--- program BumperR_C (robot ABB IRB 1300-10/1.15) ---
  Smooth(1)
  Set speed (1000.0 mm/s)
  Set Ref.: Bumper_R
  Set Tool: Generic Paint Sprayer
  Show Generic Paint Sprayer
  MoveJ 1 to (-1936.32, -807.88, 631.21) mm, rotated rx 93.18 ry 4.14 rz 127.64 deg; joints [-99.533, -17.421, 17.763, 90.671, 92.041, 174.508, 166.076, 424.987, 537.758]
  MoveL 2 to (-1936.32, -807.88, 631.21) mm, rotated rx 93.18 ry 4.14 rz 127.64 deg; joints [-99.533, -17.421, 17.763, 90.671, 92.041, 174.508, 166.076, 424.987, 537.758]
  MoveL 3 to (-1857.02, -747.22, 625.67) mm, rotated rx 93.18 ry 4.14 rz 127.64 deg; joints [-99.533, -17.421, 17.763, 90.671, 92.041, 174.508, 245.383, 485.648, 543.299]
  MoveL 4 to (-1857.02, -747.22, 625.67) mm, rotated rx 93.18 ry 4.14 rz 127.64 deg; joints [-99.533, -17.421, 17.763, 90.671, 92.041, 174.508, 245.383, 485.648, 543.299]
  Set speed (200.0 mm/s)
  MoveL 5 to (-1854.92, -751.4, 608.66) mm, rotated rx 92.71 ry 3.53 rz 127.58 deg; joints [-99.511, -17.421, 17.763, 90.568, 92.041, 175.269, 247.254, 481.589, 561.94]
  MoveL 6 to (-1853.09, -755.07, 592.18) mm, rotated rx 92.47 ry 3.35 rz 126.5 deg; joints [-99.489, -17.145, 17.763, 90.433, 93.086, 175.269, 247.254, 484.938, 580.964]
  MoveL 7 to (-1851.52, -758.47, 576.48) mm, rotated rx 93.66 ry 4.99 rz 126.32 deg; joints [-99.364, -17.145, 16.133, 90.721, 93.228, 174.897, 247.254, 485.358, 580.964]
  MoveL 8 to (-1850.74, -761.61, 561.83) mm, rotated rx 94.86 ry 6.58 rz 126.56 deg; joints [-99.364, -17.392, 14.819, 91.032, 93.106, 174.504, 247.642, 485.358, 580.964]
  MoveL 9 to (-1850.48, -763.96, 548.75) mm, rotated rx 96.79 ry 9.07 rz 127.08 deg; joints [-99.364, -17.665, 14.066, 91.464, 92.867, 172.428, 247.79, 485.358, 580.964]
  MoveL 10 to (-1851.52, -765.27, 536.72) mm, rotated rx 100.03 ry 13.16 rz 127.84 deg; joints [-99.41, -17.665, 13.808, 92.093, 92.867, 167.569, 247.288, 485.542, 580.964]
  MoveL 11 to (-1854.14, -765.79, 525.73) mm, rotated rx 106.46 ry 20.29 rz 130.44 deg; joints [-99.565, -17.69, 13.808, 93.445, 92.604, 158.33, 247.288, 485.542, 571.446]
  MoveL 12 to (-1858.59, -765.01, 515.26) mm, rotated rx 114.08 ry 25.91 rz 135.64 deg; joints [-99.582, -18.538, 13.808, 95.79, 90.846, 150.452, 247.288, 485.542, 548.94]
  MoveL 13 to (-1865.65, -762.91, 505.32) mm, rotated rx 122.27 ry 29.64 rz 141.93 deg; joints [-99.582, -19.151, 13.808, 98.838, 88.998, 143.312, 247.792, 485.542, 521.609]
  MoveL 14 to (-1874.81, -759.25, 495.64) mm, rotated rx 129.05 ry 31.24 rz 147.4 deg; joints [-99.584, -19.274, 13.808, 101.789, 87.65, 137.836, 247.792, 485.542, 499.519]
  MoveL 15 to (-1886.32, -754.02, 486.49) mm, rotated rx 136.02 ry 31.67 rz 153.13 deg; joints [-99.584, -19.274, 13.808, 105.29, 86.453, 132.536, 248.559, 488.116, 473.738]
  MoveL 16 to (-1899.66, -746.96, 478.12) mm, rotated rx 142.32 ry 31.02 rz 158.3 deg; joints [-99.584, -19.274, 13.808, 108.952, 85.547, 127.949, 249.413, 495.397, 447.495]
  MoveL 17 to (-1915.36, -738.32, 470.27) mm, rotated rx 145.68 ry 30.62 rz 160.83 deg; joints [-99.727, -19.274, 13.808, 110.865, 85.547, 125.497, 241.966, 507.62, 437.97]
  MoveL 18 to (-1931.84, -728.38, 462.94) mm, rotated rx 149.65 ry 30.54 rz 163.43 deg; joints [-99.727, -19.274, 13.808, 112.679, 85.974, 122.436, 231.514, 526.497, 429.039]
  MoveL 19 to (-1948.58, -717.13, 456.14) mm, rotated rx 152.24 ry 30.71 rz 164.95 deg; joints [-99.727, -19.274, 13.808, 113.594, 86.536, 120.405, 217.15, 545.852, 427.786]
  MoveL 20 to (-1964.28, -704.84, 450.12) mm, rotated rx 153.43 ry 32.04 rz 165.14 deg; joints [-99.727, -19.274, 12.548, 112.864, 87.093, 120.405, 195.765, 569.427, 430.366]
  MoveL 21 to (-1978.14, -692.28, 444.63) mm, rotated rx 153.62 ry 34.41 rz 164.34 deg; joints [-99.727, -19.274, 11.863, 110.908, 88.335, 120.405, 170.573, 593.858, 448.118]
  MoveL 22 to (-1990.18, -678.94, 439.66) mm, rotated rx 153.89 ry 36.46 rz 163.77 deg; joints [-99.727, -19.274, 11.132, 109.278, 89.362, 120.405, 149.601, 617.715, 462.665]
  MoveL 23 to (-2001.17, -663.76, 435.73) mm, rotated rx 154.97 ry 37.74 rz 164.05 deg; joints [-99.727, -19.274, 9.965, 108.565, 89.866, 120.405, 133.981, 642.57, 464.996]
  MoveL 24 to (-2011.11, -646.76, 432.33) mm, rotated rx 155.17 ry 39.62 rz 163.56 deg; joints [-99.727, -19.274, 9.284, 107.066, 90.789, 120.405, 116.666, 668.628, 477.923]
  MoveL 25 to (-2020.53, -627.4, 429.98) mm, rotated rx 157.04 ry 40.04 rz 164.76 deg; joints [-99.727, -19.274, 9.179, 107.28, 91.159, 119.081, 107.159, 693.484, 477.923]
  MoveL 26 to (-2029.16, -606.21, 428.41) mm, rotated rx 158.94 ry 40.39 rz 165.99 deg; joints [-99.727, -19.274, 9.179, 107.517, 91.545, 117.663, 98.62, 719.886, 477.702]
  MoveL 27 to (-2037.01, -583.97, 427.36) mm, rotated rx 160.23 ry 41.22 rz 166.67 deg; joints [-99.727, -19.274, 8.49, 107.168, 91.913, 117.224, 88.381, 748.859, 477.702]
  MoveL 28 to (-2044.59, -558.86, 426.58) mm, rotated rx 161.39 ry 42.2 rz 167.25 deg; joints [-99.727, -19.274, 7.571, 106.639, 92.277, 117.063, 77.677, 781.257, 477.702]
  MoveL 29 to (-2052.44, -527.72, 426.05) mm, rotated rx 163.85 ry 43.54 rz 168.72 deg; joints [-99.727, -19.274, 6.547, 106.072, 92.915, 116.051, 66.17, 823.308, 477.702]
  MoveL 30 to (-2059.77, -491.62, 425.27) mm, rotated rx 165.59 ry 45.05 rz 169.7 deg; joints [-99.727, -19.274, 4.995, 105.182, 93.397, 116.035, 54.117, 870.014, 477.702]
  MoveL 31 to (-2066.57, -450.02, 425.01) mm, rotated rx 167.57 ry 45.52 rz 171.06 deg; joints [-99.727, -19.274, 4.773, 105.136, 93.752, 114.842, 46.502, 916.944, 477.702]
  MoveL 32 to (-2072.32, -407.9, 424.48) mm, rotated rx 169.72 ry 45.69 rz 172.6 deg; joints [-99.727, -19.274, 4.772, 105.319, 94.067, 113.385, 40.863, 963.663, 477.247]
  MoveL 33 to (-2076.77, -369.45, 424.48) mm, rotated rx 172.37 ry 44.66 rz 174.62 deg; joints [-99.739, -19.073, 4.773, 106.624, 94.061, 111.6, 40.863, 1004.094, 466.401]
  MoveL 34 to (-2080.43, -332.3, 424.22) mm, rotated rx 173.02 ry 44.75 rz 175.07 deg; joints [-99.739, -19.073, 4.699, 106.632, 94.169, 111.22, 37.023, 1042.993, 466.401]
  MoveL 35 to (-2083.57, -293.84, 424.22) mm, rotated rx 174.33 ry 44.89 rz 175.99 deg; joints [-99.739, -19.073, 4.643, 106.655, 94.406, 110.368, 33.624, 1084.71, 466.401]
  MoveL 36 to (-2086.45, -254.34, 423.96) mm, rotated rx 174.99 ry 44.96 rz 176.45 deg; joints [-99.739, -19.073, 4.578, 106.671, 94.512, 109.977, 30.611, 1125.93, 466.401]
  MoveL 37 to (-2088.81, -213.79, 423.96) mm, rotated rx 174.99 ry 44.96 rz 176.45 deg; joints [-99.739, -19.073, 4.578, 106.671, 94.512, 109.977, 28.256, 1166.48, 466.401]
  MoveL 38 to (-2090.9, -172.19, 423.96) mm, rotated rx 176.32 ry 45.06 rz 177.39 deg; joints [-99.739, -19.073, 4.541, 106.71, 94.746, 109.105, 25.989, 1211.272, 466.401]
  MoveL 39 to (-2092.47, -129.81, 423.96) mm, rotated rx 177.06 ry 44.63 rz 177.93 deg; joints [-99.74, -19.032, 4.541, 107.175, 94.739, 108.614, 25.988, 1254.666, 462.512]
  MoveL 40 to (-2093.78, -86.9, 424.22) mm, rotated rx 178.13 ry 43.73 rz 178.71 deg; joints [-99.74, -19.032, 4.541, 108.117, 94.642, 107.976, 27.818, 1299.855, 454.042]
  MoveL 41 to (-2094.82, -43.48, 424.22) mm, rotated rx 179.06 ry 43.76 rz 179.35 deg; joints [-99.74, -19.032, 4.528, 108.161, 94.823, 107.343, 26.715, 1345.663, 454.042]
  MoveL 42 to (-2095.87, -0.05, 424.22) mm, rotated rx -180 ry 43.76 rz -180 deg; joints [-99.74, -19.031, 4.528, 108.215, 95.004, 106.699, 25.661, 1391.44, 454.042]
  MoveL 43 to (-2094.82, 43.64, 424.22) mm, rotated rx -179.06 ry 43.76 rz -179.35 deg; joints [-99.572, -19.031, 4.528, 108.223, 95.03, 106.004, 25.661, 1437.299, 454.038]
  MoveL 44 to (-2093.78, 87.07, 424.22) mm, rotated rx -178.13 ry 43.73 rz -178.71 deg; joints [-99.397, -19.031, 4.528, 108.24, 95.047, 105.308, 25.661, 1482.893, 453.951]
  MoveL 45 to (-2092.47, 129.97, 423.96) mm, rotated rx -177.06 ry 44.63 rz -177.93 deg; joints [-99.397, -19.031, 3.701, 107.472, 95.232, 105.308, 23.483, 1530.189, 456.644]
  MoveL 46 to (-2090.9, 172.35, 423.96) mm, rotated rx -176.32 ry 45.06 rz -177.39 deg; joints [-99.397, -19.031, 3.152, 107.121, 95.314, 105.308, 23.335, 1575.521, 456.873]
  MoveL 47 to (-2088.81, 213.69, 423.96) mm, rotated rx -174.99 ry 44.96 rz -176.45 deg; joints [-99.155, -19.031, 3.152, 107.158, 95.314, 104.338, 24.086, 1619.712, 456.608]
  MoveL 48 to (-2086.45, 254.24, 423.96) mm, rotated rx -174.99 ry 44.96 rz -176.45 deg; joints [-99.155, -19.031, 3.152, 107.158, 95.314, 104.338, 26.44, 1660.262, 456.608]
  MoveL 49 to (-2083.57, 293.74, 424.22) mm, rotated rx -174.33 ry 44.89 rz -175.99 deg; joints [-99.036, -19.031, 3.152, 107.184, 95.314, 103.855, 28.685, 1701.202, 456.156]
  MoveL 50 to (-2080.43, 332.2, 424.22) mm, rotated rx -173.02 ry 44.75 rz -175.07 deg; joints [-98.796, -19.031, 3.152, 107.239, 95.314, 102.892, 30.574, 1742.548, 455.762]
  MoveL 51 to (-2076.77, 369.61, 424.48) mm, rotated rx -172.55 ry 44.21 rz -174.79 deg; joints [-98.796, -19.031, 3.152, 107.761, 95.299, 102.576, 35.936, 1781.615, 451.106]
  MoveL 52 to (-2072.32, 408.07, 424.48) mm, rotated rx -169.84 ry 45.47 rz -172.72 deg; joints [-98.796, -19.031, 1.231, 106.589, 95.496, 102.576, 34.759, 1829.747, 451.505]
  MoveL 53 to (-2066.57, 450.19, 425.01) mm, rotated rx -167.57 ry 45.52 rz -171.06 deg; joints [-98.445, -19.031, 0.86, 106.319, 95.496, 101.296, 37.362, 1877.139, 451.505]
  MoveL 54 to (-2059.77, 491.52, 425.27) mm, rotated rx -165.59 ry 45.05 rz -169.7 deg; joints [-98.116, -19.031, 0.86, 106.5, 95.496, 99.832, 42.872, 1922.962, 449.946]
  MoveL 55 to (-2052.44, 527.89, 426.05) mm, rotated rx -164.03 ry 43.34 rz -168.89 deg; joints [-97.985, -19.031, 0.86, 107.995, 95.496, 98.569, 54.252, 1966.24, 436.98]
  MoveL 56 to (-2044.59, 558.76, 426.58) mm, rotated rx -161.39 ry 42.2 rz -167.25 deg; joints [-97.449, -19.031, 0.86, 108.62, 95.496, 96.434, 61.329, 2005.2, 431.733]
  MoveL 57 to (-2037.01, 584.14, 427.36) mm, rotated rx -159.73 ry 41 rz -166.38 deg; joints [-97.078, -19.031, 0.86, 109.449, 95.496, 94.99, 69.884, 2037.373, 424.494]
  MoveL 58 to (-2029.16, 606.11, 428.41) mm, rotated rx -158.46 ry 40.17 rz -165.72 deg; joints [-96.751, -19.031, 0.86, 109.96, 95.496, 93.867, 77.91, 2064.498, 419.566]
  MoveL 59 to (-2020.53, 627.3, 429.98) mm, rotated rx -157.04 ry 40.04 rz -164.76 deg; joints [-96.751, -19.031, 0.73, 109.835, 95.79, 92.944, 85.922, 2089.517, 419.566]
  MoveL 60 to (-2011.11, 646.92, 432.33) mm, rotated rx -155.42 ry 39.47 rz -163.79 deg; joints [-96.299, -19.031, 0.73, 109.921, 95.79, 91.528, 93.399, 2114.204, 416.903]
  MoveL 61 to (-2001.17, 663.93, 435.73) mm, rotated rx -155.23 ry 37.59 rz -164.28 deg; joints [-96.106, -19.031, 0.73, 111.729, 95.79, 91.025, 109.339, 2138.748, 399.131]
  MoveL 62 to (-1990.18, 678.84, 439.66) mm, rotated rx -154.15 ry 36.32 rz -163.99 deg; joints [-95.651, -19.031, 0.73, 112.633, 95.79, 89.863, 121.839, 2160.968, 388.385]
  MoveL 63 to (-1978.14, 692.44, 444.63) mm, rotated rx -153.62 ry 34.41 rz -164.34 deg; joints [-95.237, -19.031, 0.73, 114.331, 95.79, 89.028, 139.219, 2183.618, 370.37]
  MoveL 64 to (-1964.28, 705, 450.12) mm, rotated rx -153.68 ry 31.92 rz -165.34 deg; joints [-94.887, -19.031, 0.73, 116.823, 95.79, 88.593, 162.975, 2206.59, 345.904]
  MoveL 65 to (-1948.58, 717.03, 456.14) mm, rotated rx -152.24 ry 30.71 rz -164.95 deg; joints [-94.076, -19.031, 0.73, 117.431, 95.79, 86.979, 178.162, 2227.857, 335.852]
  MoveL 66 to (-1931.84, 728.28, 462.94) mm, rotated rx -149.65 ry 30.54 rz -163.43 deg; joints [-94.076, -19.031, 0.546, 116.895, 96.626, 85.113, 192.486, 2247.762, 335.852]
  MoveL 67 to (-1915.36, 738.49, 470.27) mm, rotated rx -145.68 ry 30.62 rz -160.83 deg; joints [-94.076, -19.031, -0.772, 115.634, 97.273, 83.206, 202.648, 2270.964, 335.852]
  MoveL 68 to (-1899.66, 747.12, 478.12) mm, rotated rx -142.32 ry 31.02 rz -158.3 deg; joints [-94.076, -19.031, -2.193, 114.066, 97.487, 81.93, 210.701, 2287.64, 335.852]
  MoveL 69 to (-1886.32, 753.92, 486.49) mm, rotated rx -136.33 ry 31.66 rz -153.39 deg; joints [-94.433, -19.031, -5.824, 111.213, 97.484, 80.878, 211.61, 2307.705, 336.675]
  MoveL 70 to (-1874.81, 759.15, 495.64) mm, rotated rx -129.05 ry 31.24 rz -147.4 deg; joints [-94.884, -19.031, -10.183, 108.228, 97.484, 79.328, 211.337, 2327.777, 336.675]
  MoveL 71 to (-1865.65, 762.82, 505.32) mm, rotated rx -121.95 ry 29.53 rz -141.67 deg; joints [-95.215, -19.031, -14.028, 105.588, 97.484, 76.903, 210.999, 2343.299, 336.676]
  MoveL 72 to (-1858.59, 764.91, 515.26) mm, rotated rx -113.78 ry 25.73 rz -135.42 deg; joints [-95.671, -19.031, -18.384, 102.957, 97.484, 73.021, 209.766, 2357.906, 336.68]
  MoveL 73 to (-1854.14, 765.7, 525.73) mm, rotated rx -105.9 ry 19.78 rz -130.1 deg; joints [-96.122, -19.031, -22.104, 100.789, 97.484, 67.188, 208.374, 2368.079, 336.681]
  MoveL 74 to (-1851.52, 765.43, 536.72) mm, rotated rx -100.03 ry 13.16 rz -127.84 deg; joints [-96.122, -19.031, -23.565, 99.944, 97.888, 59.882, 208.876, 2376.573, 336.681]
  MoveL 75 to (-1850.48, 763.86, 548.75) mm, rotated rx -97.28 ry 9.68 rz -127.23 deg; joints [-96.122, -19.033, -23.565, 99.613, 98.284, 55.461, 209.792, 2376.573, 333.147]
  MoveL 76 to (-1850.74, 761.51, 561.83) mm, rotated rx -94.38 ry 5.95 rz -126.45 deg; joints [-96.122, -19.324, -23.565, 99.024, 98.427, 50.977, 208.321, 2376.573, 329.103]
  MoveL 77 to (-1851.52, 758.63, 576.48) mm, rotated rx -93.66 ry 4.99 rz -126.32 deg; joints [-96.122, -19.541, -23.565, 98.92, 98.45, 49.99, 207.062, 2376.573, 316.404]
  MoveL 78 to (-1853.09, 755.23, 592.18) mm, rotated rx -92.47 ry 3.35 rz -126.5 deg; joints [-96.122, -19.581, -23.565, 98.982, 98.785, 48.026, 205.933, 2376.573, 304.255]
  MoveL 79 to (-1854.92, 751.31, 608.66) mm, rotated rx -92.71 ry 3.53 rz -127.58 deg; joints [-95.902, -19.193, -23.565, 99.595, 99.379, 48.025, 205.932, 2376.585, 287.089]
  MoveL 80 to (-1857.02, 747.38, 625.67) mm, rotated rx -92.47 ry 3.22 rz -127.55 deg; joints [-95.903, -19.46, -23.565, 99.595, 99.364, 47.903, 203.405, 2376.585, 270.462]
  Set speed (1000.0 mm/s)
  MoveL 81 to (-1857.02, 747.38, 625.67) mm, rotated rx -92.47 ry 3.22 rz -127.55 deg; joints [-95.903, -19.46, -23.565, 99.595, 99.364, 47.903, 203.405, 2376.585, 270.462]
  MoveL 82 to (-1936.37, 808.08, 629.98) mm, rotated rx -92.47 ry 3.22 rz -127.55 deg; joints [-95.903, -19.46, -23.565, 99.595, 99.364, 47.903, 124.049, 2437.282, 266.151]
  Set speed (1000.0 mm/s)
  MoveL 83 to (-1866.33, 853.74, 600.09) mm, rotated rx -83.63 ry -41.53 rz -164.5 deg; joints [-62.31, -26.599, -19.684, 114.622, 92.23, 9.806, 295.721, 2881.383, 207.551]
  MoveL 84 to (-1832.69, 759.94, 608.4) mm, rotated rx -85.23 ry -1.7 rz -160.41 deg; joints [0, -20.746, 0, 63.366, 46.167, 29.285, 22.945, 2896.284, 466.116]
  MoveL 85 to (-1832.69, 759.94, 608.4) mm, rotated rx -85.23 ry -1.7 rz -160.41 deg; joints [0, -20.746, 0, 63.366, 46.167, 29.285, 22.945, 2896.284, 466.116]
  Set speed (200.0 mm/s)
  MoveL 86 to (-1807.05, 769.62, 608.4) mm, rotated rx -85.47 ry -1.55 rz -161.18 deg; joints [0.673, -20.681, 0, 63.662, 46.168, 29.285, 53.093, 2915.113, 464.886]
  MoveL 87 to (-1774.35, 780.87, 608.4) mm, rotated rx -86.88 ry -1.04 rz -161.54 deg; joints [0.494, -20.669, 0, 65.263, 46.167, 29.285, 88.293, 2928.573, 454.825]
  MoveL 88 to (-1737.72, 792.64, 608.92) mm, rotated rx -87.13 ry -0.81 rz -164.2 deg; joints [2.732, -20.666, 0, 65.706, 46.49, 29.285, 144.085, 2970.228, 453.078]
  MoveL 89 to (-1699.52, 803.37, 611.02) mm, rotated rx -87.04 ry -0.78 rz -165.26 deg; joints [3.621, -20.666, 0, 65.706, 46.681, 29.257, 190.209, 2992.448, 451.942]
  MoveL 90 to (-1699.52, 803.37, 611.02) mm, rotated rx -87.81 ry -2 rz -137.59 deg; joints [-23.141, -21.64, 0, 65.706, 45.639, 29.257, 72.494, 2638.724, 437.476]
  MoveL 91 to (-1692.72, 808.6, 595.58) mm, rotated rx -87.36 ry -2.41 rz -137.69 deg; joints [-23.141, -21.452, 0, 65.706, 45.726, 28.553, 77.414, 2643.64, 455.753]
  MoveL 92 to (-1682.78, 815.66, 576.22) mm, rotated rx -85.22 ry -4.18 rz -138.93 deg; joints [-23.14, -21.036, 0, 65.706, 46.944, 25.645, 86.714, 2657.383, 487.623]
  MoveL 93 to (-1678.33, 821.16, 555.29) mm, rotated rx -92.02 ry 1.97 rz -135.8 deg; joints [-23.14, -21.586, 0, 66.424, 43.225, 34.246, 86.714, 2640.571, 472.908]
  MoveL 94 to (-1642.49, 837.12, 523.37) mm, rotated rx -77.29 ry -8.01 rz -148.28 deg; joints [-23.14, -19.929, 0, 66.424, 55.746, 16.427, 152.9, 2736.554, 595.298]
  MoveL 95 to (-1620.52, 847.58, 496.95) mm, rotated rx -79.58 ry -7.51 rz -144.62 deg; joints [-23.14, -19.686, 0, 66.424, 52.076, 18.199, 155.26, 2721.165, 605.579]
  MoveL 96 to (-1620.52, 847.58, 496.95) mm, rotated rx -99.89 ry 2.5 rz -165.96 deg; joints [-23.14, -12.952, 0, 92.6, 67.432, 18.199, 210.874, 2845.232, 499.77]
  MoveL 97 to (-1641.45, 845.49, 477.07) mm, rotated rx -98.6 ry 2.33 rz -164.94 deg; joints [-23.14, -13.332, 0, 91.157, 66.772, 18.199, 186.996, 2840.685, 528.15]
  MoveL 98 to (-1660.28, 843.13, 455.62) mm, rotated rx -97.18 ry 2.02 rz -164.37 deg; joints [-23.141, -13.834, 0, 89.716, 66.592, 18.199, 170.028, 2839.081, 558.046]
  MoveL 99 to (-1678.33, 840.52, 432.86) mm, rotated rx -96.24 ry 1.87 rz -163.38 deg; joints [-23.141, -14.087, 0, 88.595, 65.882, 18.199, 147.906, 2832.55, 587.081]
  MoveL 100 to (-1695.08, 837.64, 409.05) mm, rotated rx -95.06 ry 1.57 rz -162.84 deg; joints [-23.141, -14.51, 0, 87.369, 65.678, 18.199, 132.362, 2829.437, 617.84]
  MoveL 101 to (-1709.73, 835.02, 384.98) mm, rotated rx -93.88 ry 1.24 rz -162.32 deg; joints [-23.141, -14.941, 0, 86.142, 65.486, 18.199, 119.084, 2826.443, 648.781]
  MoveL 102 to (-1722.28, 832.41, 361.44) mm, rotated rx -92.94 ry 0.99 rz -161.35 deg; joints [-23.141, -15.215, 0, 85.008, 64.801, 18.199, 102.986, 2819.412, 678.238]
  MoveL 103 to (-1732.23, 830.05, 338.68) mm, rotated rx -92 ry 0.68 rz -161.32 deg; joints [-23.127, -15.625, 0, 84.119, 65.017, 18.199, 97.559, 2819.356, 706.065]
  MoveL 104 to (-1740.6, 827.96, 316.96) mm, rotated rx -91.53 ry 0.52 rz -161.31 deg; joints [-23.126, -15.833, 0, 83.678, 65.137, 18.199, 91.508, 2818.353, 730.315]
  MoveL 105 to (-1747.4, 826.13, 295.51) mm, rotated rx -91.06 ry 0.37 rz -160.6 deg; joints [-23.4, -15.978, 0, 83.118, 64.841, 18.199, 82.237, 2810.955, 754.634]
  Set speed (1000.0 mm/s)
  MoveL 106 to (-1747.4, 826.13, 295.51) mm, rotated rx -91.06 ry 0.37 rz -160.6 deg; joints [-23.4, -15.978, 0, 83.118, 64.841, 18.199, 82.237, 2810.955, 754.634]
  MoveL 107 to (-1780.63, 920.43, 297.36) mm, rotated rx -91.06 ry 0.37 rz -160.6 deg; joints [-23.4, -15.978, 0, 83.118, 64.841, 18.199, 49.007, 2905.255, 752.786]
  Set speed (1000.0 mm/s)
  MoveL 108 to (-1840, 893.27, 313.81) mm, rotated rx -106.34 ry 6.01 rz -160.35 deg; joints [-23.4, -17.541, 0, 92.672, 59.812, 27.622, 0.008, 2861.075, 623.578]
  MoveL 109 to (-1804.95, 803.89, 285.83) mm, rotated rx -106.34 ry 6.01 rz -160.35 deg; joints [-23.4, -17.541, 0, 92.672, 59.812, 27.622, 35.053, 2771.694, 651.559]
  MoveL 110 to (-1804.95, 803.89, 285.83) mm, rotated rx -106.34 ry 6.01 rz -160.35 deg; joints [-23.4, -17.541, 0, 92.672, 59.812, 27.622, 35.053, 2771.694, 651.559]
  Set speed (200.0 mm/s)
  MoveL 111 to (-1832.95, 791.59, 290.54) mm, rotated rx -106.49 ry 6.19 rz -159.99 deg; joints [-23.4, -17.541, 0.133, 92.672, 59.412, 27.666, 4.112, 2756.326, 647.26]
  MoveL 112 to (-1858.06, 779.82, 294.2) mm, rotated rx -106.41 ry 7.21 rz -156.92 deg; joints [-26.51, -20.886, 1.667, 90.881, 59.412, 30.95, 0, 2721.012, 647.26]
  MoveL 113 to (-1879.78, 768.57, 296.56) mm, rotated rx -105.99 ry 7.97 rz -154.18 deg; joints [-29.001, -23.988, 2.357, 88.525, 59.412, 34.604, 0, 2695.317, 647.26]
  MoveL 114 to (-1896.78, 758.89, 298.13) mm, rotated rx -106.1 ry 9.48 rz -150.31 deg; joints [-32.699, -26.95, 2.767, 86.07, 59.412, 39.328, 0, 2657.479, 647.26]
  MoveL 115 to (-1911.69, 749.48, 299.17) mm, rotated rx -106.56 ry 10.61 rz -148.24 deg; joints [-34.777, -29.185, 3.342, 84.726, 59.412, 42.61, 0, 2636.415, 647.26]
  MoveL 116 to (-1927.13, 738.75, 299.96) mm, rotated rx -105.67 ry 11.02 rz -145.73 deg; joints [-36.306, -31.519, 3.342, 81.953, 59.412, 45.771, 0, 2619.867, 652.638]
  MoveL 117 to (-1942.56, 726.98, 301) mm, rotated rx -105.75 ry 12.18 rz -143.21 deg; joints [-38.217, -33.858, 3.342, 79.586, 59.412, 49.888, 0, 2598.73, 654.329]
  MoveL 118 to (-1957.74, 714.42, 301.79) mm, rotated rx -105.83 ry 13.67 rz -140.19 deg; joints [-40.307, -36.353, 3.342, 76.719, 59.412, 54.629, 0, 2574.299, 659.016]
  MoveL 119 to (-1971.86, 701.08, 302.57) mm, rotated rx -105.19 ry 14.87 rz -136.61 deg; joints [-42.079, -38.903, 3.342, 72.981, 59.412, 59.147, 0, 2548.829, 669.678]
  MoveL 120 to (-1984.68, 686.95, 303.1) mm, rotated rx -104.58 ry 16.89 rz -131.85 deg; joints [-44.246, -41.542, 3.342, 68.194, 59.412, 64.909, 0, 2512.396, 685.44]
  MoveL 121 to (-1996.19, 672.3, 303.62) mm, rotated rx -105.37 ry 20.17 rz -128.56 deg; joints [-45.598, -43.63, 3.342, 64.184, 59.412, 71.634, 0, 2480.166, 696.443]
  MoveL 122 to (-2006.4, 656.6, 303.88) mm, rotated rx -105.16 ry 23.11 rz -124.63 deg; joints [-46.174, -45.488, 3.342, 58.938, 59.412, 77.967, 0, 2443.432, 714.605]
  MoveL 123 to (-2015.55, 640.12, 304.14) mm, rotated rx -105.39 ry 26.98 rz -121.25 deg; joints [-46.174, -47.75, 3.343, 53.282, 60.14, 85.802, 7.235, 2413.258, 735.61]
  MoveL 124 to (-2023.66, 622.59, 304.14) mm, rotated rx -105.02 ry 30.09 rz -118.16 deg; joints [-46.174, -47.998, 3.343, 49.217, 60.37, 90.526, 0.63, 2370.196, 753.089]
  MoveL 125 to (-2030.47, 604.8, 304.14) mm, rotated rx -104.12 ry 31.18 rz -115.91 deg; joints [-46.181, -48.648, 3.343, 46.493, 60.949, 92.894, 0.01, 2341.413, 766.26]
  MoveL 126 to (-2036.48, 586.75, 303.88) mm, rotated rx -103.81 ry 32.8 rz -114.41 deg; joints [-46.851, -49.255, 3.343, 45.076, 62.033, 95.231, 0, 2316.688, 777.689]
  MoveL 127 to (-2041.98, 569.22, 303.88) mm, rotated rx -105.4 ry 36.74 rz -114.72 deg; joints [-46.853, -49.837, 3.343, 44.146, 63.26, 100.087, 0, 2300.801, 786.26]
  MoveL 128 to (-2046.42, 552.48, 303.62) mm, rotated rx -106.11 ry 42.57 rz -113.12 deg; joints [-47.479, -50.038, 3.343, 41.986, 65.443, 106.494, 0, 2270.786, 809.046]
  MoveL 129 to (-2050.61, 534.69, 303.62) mm, rotated rx -109.1 ry 48.54 rz -114.8 deg; joints [-47.479, -50.429, 3.343, 41.714, 67.353, 112.969, 0, 2258.639, 820.752]
  MoveL 130 to (-2054.53, 514.02, 303.36) mm, rotated rx -110.56 ry 52.74 rz -115.23 deg; joints [-47.479, -50.69, 3.343, 40.989, 68.994, 117.465, 0, 2238.905, 834.382]
  MoveL 131 to (-2058.2, 490.48, 303.88) mm, rotated rx -114 ry 59.08 rz -117.43 deg; joints [-47.479, -50.872, 3.343, 40.753, 71.292, 123.95, 0, 2220.446, 850.258]
  MoveL 132 to (-2061.08, 464.84, 305.97) mm, rotated rx -122.64 ry 66.68 rz -124.9 deg; joints [-47.479, -51.083, 3.343, 41.781, 73.743, 131.949, 0, 2208.96, 860.36]
  MoveL 133 to (-2062.65, 439.2, 310.16) mm, rotated rx -130.58 ry 72.26 rz -131.97 deg; joints [-47.479, -50.951, 3.343, 42.168, 75.885, 137.566, 0.014, 2190.405, 870.985]
  MoveL 134 to (-2062.91, 416.18, 317.48) mm, rotated rx -143.56 ry 74.86 rz -144.52 deg; joints [-47.479, -51.111, 3.343, 43.565, 76.5, 141.58, 0.003, 2178.849, 861.295]
  MoveL 135 to (-2061.86, 396.56, 326.64) mm, rotated rx -154.06 ry 77.62 rz -154.59 deg; joints [-47.479, -50.7, 3.343, 43.858, 77.758, 144.603, 0.003, 2161.713, 861.88]
  MoveL 136 to (-2060.55, 380.6, 335.8) mm, rotated rx 150.62 ry 75.7 rz 151.38 deg; joints [-45.847, -50.793, 3.343, 46.572, 77.758, 156.331, 0, 2171.642, 840.226]
  MoveL 137 to (-2058.72, 368.04, 344.43) mm, rotated rx 152.54 ry 74.9 rz 153.36 deg; joints [-45.847, -50.981, 3.343, 46.912, 77.016, 156.331, 1.624, 2159.565, 823.551]
  MoveL 138 to (-2058.72, 368.04, 344.43) mm, rotated rx 92.19 ry 15.16 rz 98.34 deg; joints [-44.513, -50.981, 6.874, 68.618, 77.016, 213.54, 0.029, 2281.819, 776.099]
  MoveL 139 to (-2057.15, 355.75, 333.7) mm, rotated rx 92.56 ry 14.93 rz 99.84 deg; joints [-45.621, -51.277, 6.873, 68.618, 76.619, 213.86, 0.028, 2259.663, 783.809]
  MoveL 140 to (-2055.32, 342.93, 324.29) mm, rotated rx 92.93 ry 15.77 rz 100.68 deg; joints [-45.895, -51.277, 6.089, 67.95, 76.619, 213.86, 3.03, 2242.747, 789.664]
  MoveL 141 to (-2053.23, 328.54, 316.96) mm, rotated rx 95.76 ry 28.51 rz 101.93 deg; joints [-45.895, -51.277, 6.089, 63.921, 78.506, 202.475, 4.666, 2215.059, 824.396]
  MoveL 142 to (-2051.13, 313.1, 310.68) mm, rotated rx 118.95 ry 67.19 rz 120.96 deg; joints [-45.895, -51.277, 6.033, 50.461, 78.558, 166.142, 4.666, 2125.247, 882.217]
  MoveL 143 to (-2051.92, 299.5, 309.11) mm, rotated rx -151.61 ry 73.09 rz -152.65 deg; joints [-47.318, -58.551, 5.026, 44.393, 78.558, 146.287, 59.413, 2125.246, 882.217]
  MoveL 144 to (-2052.7, 288.51, 308.07) mm, rotated rx -151.22 ry 73.16 rz -152.27 deg; joints [-47.318, -58.551, 4.959, 44.303, 78.693, 146.287, 59.104, 2114.315, 884.068]
  MoveL 145 to (-2053.49, 274.38, 306.76) mm, rotated rx -150.44 ry 73.3 rz -151.48 deg; joints [-47.318, -58.551, 4.866, 44.129, 78.934, 146.254, 59.104, 2100.102, 887.137]
  MoveL 146 to (-2054.27, 258.16, 305.97) mm, rotated rx -149.06 ry 72.23 rz -150.28 deg; joints [-47.226, -59.65, 4.866, 44.129, 78.934, 146.178, 65.904, 2092.744, 886.105]
  MoveL 147 to (-2055.06, 239.33, 305.45) mm, rotated rx -154.8 ry 72.39 rz -155.84 deg; joints [-47.225, -59.873, 4.866, 44.801, 78.77, 147.78, 65.904, 2079.049, 882.098]
  MoveL 148 to (-2056.1, 217.35, 304.93) mm, rotated rx -154.8 ry 72.39 rz -155.84 deg; joints [-47.225, -59.873, 4.866, 44.801, 78.77, 147.78, 64.858, 2057.074, 882.621]
  MoveL 149 to (-2057.15, 191.19, 304.67) mm, rotated rx -160.37 ry 72.86 rz -161.18 deg; joints [-47.225, -59.873, 4.866, 45.256, 78.83, 149.358, 63.555, 2033.518, 881.475]
  MoveL 150 to (-2057.94, 160.84, 304.4) mm, rotated rx -161.41 ry 72.47 rz -162.22 deg; joints [-47.225, -60.055, 4.866, 45.508, 78.575, 149.604, 63.555, 2005.37, 878.309]
  MoveL 151 to (-2058.98, 125, 304.14) mm, rotated rx -165.69 ry 73.35 rz -166.27 deg; joints [-47.225, -60.055, 4.866, 45.553, 79.185, 151.005, 63.203, 1971.107, 883.479]
  MoveL 152 to (-2060.03, 85.5, 303.62) mm, rotated rx -171.28 ry 73.69 rz -171.62 deg; joints [-47.225, -60.055, 4.866, 45.887, 79.393, 152.515, 62.195, 1933.866, 884.39]
  MoveL 153 to (-2060.81, 43.38, 303.36) mm, rotated rx -171.76 ry 73.23 rz -172.11 deg; joints [-47.225, -60.238, 4.866, 46.098, 79.111, 152.676, 62.196, 1893.577, 881.184]
  MoveL 154 to (-2061.6, -0.05, 302.83) mm, rotated rx -180 ry 73.41 rz -180 deg; joints [-47.225, -60.238, 4.866, 46.593, 79.366, 154.887, 61.429, 1853.309, 881.898]
  MoveL 155 to (-2060.81, -43.48, 303.36) mm, rotated rx 171.76 ry 73.23 rz 172.11 deg; joints [-47.225, -60.238, 5.04, 47.132, 79.458, 156.967, 61.428, 1812.212, 881.819]
  MoveL 156 to (-2060.03, -85.6, 303.62) mm, rotated rx 171.28 ry 73.69 rz 171.62 deg; joints [-47.225, -60.101, 5.04, 46.98, 79.805, 156.967, 61.793, 1769.226, 885.263]
  MoveL 157 to (-2058.98, -125.1, 304.14) mm, rotated rx 165.69 ry 73.35 rz 166.27 deg; joints [-47.225, -60.101, 5.219, 47.378, 79.805, 158.339, 62.013, 1731.134, 885.013]
  MoveL 158 to (-2057.94, -160.68, 304.4) mm, rotated rx 161.41 ry 72.47 rz 162.22 deg; joints [-47.225, -60.101, 5.219, 47.887, 79.452, 159.658, 62.365, 1697.132, 879.843]
  MoveL 159 to (-2057.15, -191.29, 304.67) mm, rotated rx 160.37 ry 72.86 rz 161.18 deg; joints [-47.226, -59.919, 5.219, 47.785, 79.783, 159.711, 62.365, 1665.648, 883.012]
  MoveL 160 to (-2056.1, -217.19, 304.93) mm, rotated rx 154.8 ry 72.39 rz 155.84 deg; joints [-47.226, -59.752, 5.219, 48.14, 79.98, 161.192, 62.365, 1640.946, 883.332]
  MoveL 161 to (-2055.06, -239.43, 305.45) mm, rotated rx 154.8 ry 72.39 rz 155.84 deg; joints [-47.226, -59.752, 5.219, 48.14, 79.98, 161.192, 63.412, 1618.709, 882.809]
  MoveL 162 to (-2054.27, -258.26, 305.97) mm, rotated rx 152.72 ry 72.87 rz 153.77 deg; joints [-47.226, -59.519, 5.219, 48.028, 80.515, 161.387, 63.412, 1599.29, 887.548]
  MoveL 163 to (-2053.49, -274.22, 306.76) mm, rotated rx 150.44 ry 73.3 rz 151.48 deg; joints [-47.226, -59.276, 5.219, 47.93, 81.047, 161.602, 63.411, 1582.795, 891.949]
  MoveL 164 to (-2052.7, -288.35, 308.07) mm, rotated rx 151.22 ry 73.16 rz 152.27 deg; joints [-47.226, -59.456, 5.219, 47.949, 80.936, 161.602, 65.231, 1569.676, 889.402]
  MoveL 165 to (-2051.92, -299.6, 309.11) mm, rotated rx 151.61 ry 73.09 rz 152.65 deg; joints [-47.226, -59.545, 5.22, 47.959, 80.879, 161.602, 66.522, 1558.921, 887.728]
  MoveL 166 to (-2051.13, -313.2, 310.68) mm, rotated rx -118.95 ry 67.19 rz -120.96 deg; joints [-47.226, -59.545, 3.668, 39.125, 80.879, 137.414, 80.668, 1497.992, 906.158]
  MoveL 167 to (-2053.23, -328.37, 316.96) mm, rotated rx -95.76 ry 28.51 rz -101.93 deg; joints [-56.122, -67.736, 3.668, 39.125, 79.051, 101.379, 115.031, 1497.993, 896.231]
  MoveL 168 to (-2055.32, -343.02, 324.29) mm, rotated rx -92.93 ry 15.77 rz -100.68 deg; joints [-57.194, -70.603, 3.668, 39.125, 77.241, 90.761, 126.243, 1497.993, 881.392]
  MoveL 169 to (-2057.15, -355.84, 333.7) mm, rotated rx -92.56 ry 14.93 rz -99.84 deg; joints [-57.586, -70.866, 3.668, 38.68, 77.241, 90.147, 126.243, 1481.061, 873.698]
  MoveL 170 to (-2058.72, -367.88, 344.43) mm, rotated rx -92.19 ry 15.16 rz -98.34 deg; joints [-58.148, -70.866, 3.668, 37.748, 77.445, 90.454, 126.243, 1457.761, 866.87]
  MoveL 171 to (-2058.72, -367.88, 344.43) mm, rotated rx -150.15 ry 74.39 rz -151.07 deg; joints [-40.893, -60.028, 5.104, 37.748, 78.328, 150.487, 76.801, 1457.761, 866.87]
  MoveL 172 to (-2060.55, -380.7, 335.8) mm, rotated rx 147.84 ry 77.3 rz 148.47 deg; joints [-40.893, -57.863, 5.104, 40.952, 80.981, 162.299, 61.805, 1457.762, 891.266]
  MoveL 173 to (-2061.86, -396.39, 326.64) mm, rotated rx 117.87 ry 68.52 rz 119.6 deg; joints [-40.761, -56.331, 5.215, 44.915, 80.981, 172.099, 47.4, 1457.762, 891.266]
  MoveL 174 to (-2062.91, -416.28, 317.48) mm, rotated rx 109.62 ry 57.45 rz 112.93 deg; joints [-40.761, -56.748, 5.215, 48.696, 79.77, 182.716, 46.385, 1457.762, 877.678]
  MoveL 175 to (-2062.65, -439.3, 310.16) mm, rotated rx 107.5 ry 53.36 rz 111.45 deg; joints [-40.761, -56.834, 5.215, 49.946, 79.216, 186.595, 46.385, 1440.117, 876.795]
  MoveL 176 to (-2061.08, -464.94, 305.97) mm, rotated rx 110.68 ry 54.2 rz 114.95 deg; joints [-41.782, -58.512, 5.114, 49.946, 79.216, 186.242, 58.772, 1418.26, 876.795]
  MoveL 177 to (-2058.2, -490.57, 303.88) mm, rotated rx 108.74 ry 49.93 rz 113.9 deg; joints [-41.782, -58.512, 5.114, 50.99, 78.223, 190.266, 60.275, 1393.992, 868.366]
  MoveL 178 to (-2054.53, -514.12, 303.36) mm, rotated rx 108.2 ry 47.11 rz 114.17 deg; joints [-41.782, -58.512, 5.114, 51.451, 77.052, 192.806, 62.36, 1367.394, 858.646]
  MoveL 179 to (-2050.61, -534.79, 303.62) mm, rotated rx 107.69 ry 44.45 rz 114.49 deg; joints [-41.782, -58.512, 5.114, 51.782, 75.904, 195.225, 64.918, 1342.818, 848.878]
  MoveL 180 to (-2046.42, -552.58, 303.62) mm, rotated rx 105.37 ry 39.37 rz 113.43 deg; joints [-41.782, -58.512, 5.115, 52.7, 74.899, 200.218, 68.293, 1324.841, 839.862]
  MoveL 181 to (-2041.98, -569.06, 303.88) mm, rotated rx 110.31 ry 38.82 rz 120.57 deg; joints [-44.654, -60.548, 5.115, 52.7, 72.427, 200.218, 81.675, 1290.733, 815.564]
  Set speed (1000.0 mm/s)
  MoveL 182 to (-2041.98, -569.06, 303.88) mm, rotated rx 110.31 ry 38.82 rz 120.57 deg; joints [-44.654, -60.548, 5.115, 52.7, 72.427, 200.218, 81.675, 1290.733, 815.564]
  MoveL 183 to (-2133.79, -598.01, 330.93) mm, rotated rx 110.31 ry 38.82 rz 120.57 deg; joints [-44.654, -61.802, 5.115, 52.392, 73.19, 201.26, 0.012, 1271.811, 795.076]
  Set speed (1000.0 mm/s)
  MoveL 184 to (-2128.99, -596.56, 338.03) mm, rotated rx 131.63 ry 46.89 rz 140.6 deg; joints [-48.864, -65.943, 5.115, 52.392, 69.438, 188.007, 30.804, 1271.811, 744.814]
  MoveL 185 to (-2044.07, -569.58, 292.63) mm, rotated rx 131.63 ry 46.89 rz 140.6 deg; joints [-48.864, -65.943, 5.115, 52.392, 69.438, 188.007, 115.723, 1298.788, 790.214]
  MoveL 186 to (-2044.07, -569.58, 292.63) mm, rotated rx 131.63 ry 46.89 rz 140.6 deg; joints [-48.864, -65.943, 5.115, 52.392, 69.438, 188.007, 115.723, 1298.788, 790.214]
  Set speed (200.0 mm/s)
  MoveL 187 to (-2039.1, -586.85, 292.89) mm, rotated rx 131.15 ry 44.42 rz 141.31 deg; joints [-49.298, -65.943, 5.115, 52.392, 67.641, 189.836, 122.224, 1270.616, 775.253]
  MoveL 188 to (-2033.08, -604.9, 292.89) mm, rotated rx 129.35 ry 42.65 rz 140.43 deg; joints [-49.601, -65.943, 5.115, 52.392, 67.14, 191.981, 128.459, 1247.078, 771.964]
  MoveL 189 to (-2026.28, -622.69, 292.89) mm, rotated rx 124.93 ry 37.98 rz 138.62 deg; joints [-50.632, -65.943, 5.115, 52.392, 66.012, 197.63, 135.479, 1214.12, 765.262]
  MoveL 190 to (-2018.17, -640.22, 292.89) mm, rotated rx 122.72 ry 33.45 rz 139.38 deg; joints [-52.356, -65.943, 5.115, 52.392, 64.022, 202.087, 145.312, 1174.691, 750.849]
  MoveL 191 to (-2009.28, -656.7, 292.63) mm, rotated rx 121.6 ry 29.24 rz 141.55 deg; joints [-54.713, -65.943, 5.115, 52.392, 61.721, 205.759, 157.732, 1131.841, 733.872]
  MoveL 192 to (-1998.81, -672.66, 292.37) mm, rotated rx 120.13 ry 26.12 rz 142.81 deg; joints [-56.723, -65.943, 5.115, 52.392, 60.558, 208.934, 170.482, 1096.449, 726.431]
  MoveL 193 to (-1987.3, -687.57, 291.85) mm, rotated rx 118.68 ry 21.77 rz 145.87 deg; joints [-60.383, -65.943, 5.116, 52.392, 58.628, 213.052, 188.009, 1048.513, 713.651]
  MoveL 194 to (-1974.48, -701.7, 291.32) mm, rotated rx 117.52 ry 18.52 rz 148.62 deg; joints [-63.721, -65.943, 5.116, 52.392, 57.354, 216.237, 207.019, 1006.868, 705.888]
  MoveL 195 to (-1960.09, -715.3, 290.54) mm, rotated rx 116.83 ry 16.94 rz 150.06 deg; joints [-65.544, -65.943, 5.116, 52.392, 56.863, 217.893, 224.828, 979.133, 703.837]
  MoveL 196 to (-1944.66, -728.12, 289.75) mm, rotated rx 116.46 ry 15.72 rz 151.44 deg; joints [-67.112, -65.945, 5.12, 52.392, 56.36, 219.06, 243.933, 954.254, 701.378]
  MoveL 197 to (-1928.96, -739.89, 288.97) mm, rotated rx 115.75 ry 14.06 rz 153.27 deg; joints [-69.501, -66.246, 5.12, 52.392, 56.117, 221.035, 265.227, 929.319, 701.358]
  MoveL 198 to (-1913.26, -750.62, 287.92) mm, rotated rx 115.11 ry 12.73 rz 154.82 deg; joints [-71.473, -66.302, 5.12, 52.392, 55.856, 222.542, 285.279, 905.487, 701.354]
  MoveL 199 to (-1898.35, -760.04, 286.88) mm, rotated rx 114.06 ry 10.43 rz 157.92 deg; joints [-75.322, -66.537, 5.12, 52.392, 55.503, 225.212, 309.712, 873.175, 701.354]
  MoveL 200 to (-1881.35, -769.72, 285.57) mm, rotated rx 113.93 ry 9.11 rz 160.37 deg; joints [-78.111, -67.106, 5.12, 52.392, 55.253, 226.793, 335.553, 852.932, 701.353]
  MoveL 201 to (-1859.89, -780.7, 283.47) mm, rotated rx 113.66 ry 8.41 rz 161.55 deg; joints [-79.452, -67.106, 5.12, 52.392, 55.055, 227.521, 360.987, 833.342, 702.389]
  MoveL 202 to (-1834.52, -792.48, 280.34) mm, rotated rx 112.08 ry 6.93 rz 163.44 deg; joints [-82.021, -66.469, 5.12, 52.392, 55.055, 229.262, 391.621, 797.112, 707.487]
  MoveL 203 to (-1806, -804.51, 276.15) mm, rotated rx 111.67 ry 6.7 rz 163.63 deg; joints [-82.323, -66.18, 5.12, 52.392, 55.055, 229.49, 420.465, 779.338, 712.148]
  Set speed (1000.0 mm/s)
  MoveL 204 to (-1806, -804.51, 276.15) mm, rotated rx 111.67 ry 6.7 rz 163.63 deg; joints [-82.323, -66.18, 5.12, 52.392, 55.055, 229.49, 420.465, 779.338, 712.148]
  MoveL 205 to (-1836.32, -892.47, 312.82) mm, rotated rx 111.67 ry 6.7 rz 163.63 deg; joints [-82.323, -66.18, 5.12, 52.392, 55.055, 229.49, 390.142, 691.384, 675.48]
  Set speed (1000.0 mm/s)
  MoveL 206 to (-1923.75, -805.14, 336.19) mm, rotated rx 118.21 ry 60.32 rz 121.7 deg; joints [-47.684, -66.18, 5.12, 52.392, 85.879, 183.446, 244.281, 1136.485, 887.918]
  MoveL 207 to (-1827.19, -793.79, 312.78) mm, rotated rx 118.21 ry 60.32 rz 121.7 deg; joints [-47.684, -66.18, 5.12, 52.392, 85.878, 183.446, 340.836, 1147.839, 911.328]
  MoveL 208 to (-1827.19, -793.79, 312.78) mm, rotated rx 118.21 ry 60.32 rz 121.7 deg; joints [-47.684, -66.18, 5.12, 52.392, 85.878, 183.446, 340.836, 1147.839, 911.328]
  Set speed (200.0 mm/s)
  MoveL 209 to (-1821.44, -795.88, 335.27) mm, rotated rx 121.01 ry 62.14 rz 124.22 deg; joints [-47.685, -66.391, 5.12, 51.793, 85.878, 181.469, 347.895, 1143.614, 890.319]
  MoveL 210 to (-1814.9, -797.97, 358.3) mm, rotated rx 127.49 ry 63.58 rz 130.58 deg; joints [-48.562, -67.56, 5.12, 51.793, 85.343, 179.337, 358.15, 1143.614, 862.535]
  MoveL 211 to (-1807.31, -799.8, 382.1) mm, rotated rx 131.6 ry 63.95 rz 134.66 deg; joints [-48.953, -68.335, 5.12, 51.793, 84.798, 178.4, 368.646, 1143.614, 834.182]
  Set speed (1000.0 mm/s)
  MoveL 212 to (-1807.31, -799.8, 382.1) mm, rotated rx 131.6 ry 63.95 rz 134.66 deg; joints [-48.953, -68.335, 5.12, 51.793, 84.798, 178.4, 368.646, 1143.614, 834.182]
  MoveL 213 to (-1902.42, -809.94, 411.27) mm, rotated rx 131.6 ry 63.95 rz 134.66 deg; joints [-48.953, -68.335, 5.12, 51.793, 84.798, 178.4, 273.532, 1133.474, 805.021]
  Set speed (1000.0 mm/s)
  MoveL 214 to (-1847.67, -880.23, 317.42) mm, rotated rx 99.15 ry 10.51 rz 131.44 deg; joints [-57.928, -68.335, 5.12, 51.793, 69.954, 235.57, 316.536, 919.555, 803.23]
  MoveL 215 to (-1771.73, -817.07, 301.79) mm, rotated rx 99.15 ry 10.51 rz 131.44 deg; joints [-57.928, -68.335, 5.119, 51.793, 69.954, 235.57, 392.47, 982.717, 818.856]
  MoveL 216 to (-1771.73, -817.07, 301.79) mm, rotated rx 99.15 ry 10.51 rz 131.44 deg; joints [-57.928, -68.335, 5.119, 51.793, 69.954, 235.57, 392.47, 982.717, 818.856]
  Set speed (200.0 mm/s)
  MoveL 217 to (-1765.45, -818.9, 323.5) mm, rotated rx 100.09 ry 11.62 rz 131.46 deg; joints [-57.928, -68.335, 5.119, 52.093, 69.829, 234.044, 398.343, 983.221, 793.896]
  MoveL 218 to (-1758.13, -820.99, 345.74) mm, rotated rx 102.11 ry 13.31 rz 132.99 deg; joints [-58.849, -69.231, 5.119, 52.093, 69.625, 232.228, 410.477, 983.221, 768.135]
  MoveL 219 to (-1748.97, -823.09, 368.76) mm, rotated rx 104.68 ry 15.01 rz 135.32 deg; joints [-60.299, -70.502, 5.119, 52.092, 69.27, 230.392, 426.235, 983.221, 740.437]
  MoveL 220 to (-1737.98, -825.44, 392.57) mm, rotated rx 106.79 ry 16.24 rz 137.17 deg; joints [-61.322, -71.481, 5.119, 52.092, 68.878, 228.959, 442.487, 983.221, 712.211]
  MoveL 221 to (-1724.9, -827.79, 416.9) mm, rotated rx 109.98 ry 17.71 rz 140.09 deg; joints [-62.815, -72.806, 5.119, 52.092, 68.025, 226.96, 463.176, 983.221, 679.334]
  MoveL 222 to (-1709.99, -829.89, 440.97) mm, rotated rx 111.71 ry 18.59 rz 141.31 deg; joints [-63.158, -73.283, 5.119, 52.092, 67.493, 225.612, 481.599, 983.221, 649.813]
  MoveL 223 to (-1694.03, -832.24, 464.25) mm, rotated rx 114.33 ry 19 rz 144.24 deg; joints [-64.87, -74.669, 5.119, 52.092, 66.633, 224.791, 505.193, 983.221, 619.44]
  MoveL 224 to (-1677.55, -834.07, 486.23) mm, rotated rx 116.91 ry 19.55 rz 146.6 deg; joints [-65.816, -75.5, 5.119, 52.092, 65.555, 223.398, 527.986, 983.221, 587.818]
  MoveL 225 to (-1658.97, -835.64, 507.15) mm, rotated rx 119.52 ry 19.52 rz 149.46 deg; joints [-67.31, -76.6, 5.119, 52.092, 64.311, 222.603, 554.207, 983.221, 556.814]
  MoveL 226 to (-1658.97, -835.64, 507.15) mm, rotated rx 119.33 ry -3.93 rz -173.04 deg; joints [-114.101, -88.1, 5.119, 52.092, 58.313, 251.774, 581.026, 839.271, 556.814]
  MoveL 227 to (-1687.23, -822.82, 535.15) mm, rotated rx 122.17 ry -3.34 rz -174.71 deg; joints [-112.588, -90.771, 5.119, 52.092, 57.962, 251.774, 539.405, 892.064, 536.707]
  MoveL 228 to (-1730.4, -805.82, 558.17) mm, rotated rx 127.25 ry -0.31 rz -179.59 deg; joints [-106.503, -94.719, 5.119, 52.092, 57.962, 249.108, 481.037, 991.728, 530.485]
  Set speed (1000.0 mm/s)
  MoveL 229 to (-1730.4, -805.82, 558.17) mm, rotated rx 127.25 ry -0.31 rz -179.59 deg; joints [-106.503, -94.719, 5.119, 52.092, 57.962, 249.108, 481.037, 991.728, 530.485]
  MoveL 230 to (-1729.51, -885.42, 618.69) mm, rotated rx 127.25 ry -0.31 rz -179.59 deg; joints [-106.503, -94.719, 5.12, 52.092, 57.962, 249.108, 481.925, 912.127, 469.964]
  Set speed (1000.0 mm/s)
  MoveL 231 to (-1756.3, -883.87, 638.08) mm, rotated rx 116.98 ry 5.91 rz 168.57 deg; joints [-94.276, -90.161, 5.12, 52.092, 67.067, 246.296, 445.64, 912.127, 503.708]
  MoveL 232 to (-1734.06, -797.45, 592.96) mm, rotated rx 116.98 ry 5.91 rz 168.57 deg; joints [-94.276, -90.161, 5.12, 52.092, 67.067, 246.296, 467.879, 998.555, 548.828]
  MoveL 233 to (-1734.06, -797.45, 592.96) mm, rotated rx 116.98 ry 5.91 rz 168.57 deg; joints [-94.276, -90.161, 5.12, 52.092, 67.067, 246.296, 467.879, 998.555, 548.828]
  Set speed (200.0 mm/s)
  MoveL 234 to (-1772.25, -785.41, 592.18) mm, rotated rx 117.39 ry 8.06 rz 164.86 deg; joints [-89.658, -89.452, 5.12, 52.092, 67.523, 243.612, 433.11, 1032.269, 548.828]
  MoveL 235 to (-1805.22, -773.64, 592.18) mm, rotated rx 116.25 ry 8.47 rz 163.37 deg; joints [-88.22, -88.393, 5.12, 52.092, 68.007, 243.112, 400.074, 1041.014, 548.828]
  Set speed (1000.0 mm/s)
  MoveL 236 to (-1805.22, -773.64, 592.18) mm, rotated rx 116.25 ry 8.47 rz 163.37 deg; joints [-88.22, -88.393, 5.12, 52.092, 68.007, 243.112, 400.074, 1041.014, 548.828]
  MoveL 237 to (-1837.12, -857.72, 635.92) mm, rotated rx 116.25 ry 8.47 rz 163.37 deg; joints [-88.22, -88.393, 5.12, 52.092, 68.008, 243.112, 368.169, 956.938, 505.087]
  Set speed (1000.0 mm/s)
  MoveL 238 to (-1695.61, -941.83, 266.15) mm, rotated rx 107.53 ry 4.62 rz 165.7 deg; joints [-92.114, -80.605, 5.12, 52.092, 68.008, 245.28, 509.353, 761.166, 854.867]
  MoveL 239 to (-1669.7, -850.03, 236.12) mm, rotated rx 107.53 ry 4.62 rz 165.7 deg; joints [-92.114, -80.605, 5.12, 52.092, 68.008, 245.28, 535.259, 852.966, 884.892]
  MoveL 240 to (-1669.7, -850.03, 236.12) mm, rotated rx 107.53 ry 4.62 rz 165.7 deg; joints [-92.114, -80.605, 5.12, 52.092, 68.008, 245.28, 535.259, 852.966, 884.892]
  Set speed (200.0 mm/s)
  MoveL 241 to (-1716.01, -837.21, 237.69) mm, rotated rx 110.13 ry 5.19 rz 166.14 deg; joints [-92.114, -82.886, 5.12, 51.978, 67.605, 245.116, 489.943, 890.976, 884.89]
  MoveL 242 to (-1760.74, -823.87, 239.26) mm, rotated rx 110.6 ry 5.48 rz 165.74 deg; joints [-91.608, -83.238, 5.12, 51.978, 67.605, 244.874, 444.916, 911.512, 884.004]
  MoveL 243 to (-1802.6, -810.27, 240.83) mm, rotated rx 113.25 ry 6.67 rz 164.87 deg; joints [-90.126, -85.125, 5.12, 51.978, 67.299, 243.806, 403.708, 956.144, 884.004]
  MoveL 244 to (-1838.97, -796.92, 242.4) mm, rotated rx 114.25 ry 7.88 rz 163.07 deg; joints [-87.781, -85.337, 5.12, 51.978, 67.299, 242.344, 368.41, 987.022, 881.897]
  MoveL 245 to (-1866.7, -784.89, 243.45) mm, rotated rx 115.07 ry 9.33 rz 160.88 deg; joints [-85.003, -85.337, 5.12, 51.978, 67.463, 240.622, 342.219, 1016.864, 880.954]
  MoveL 246 to (-1888.15, -774.43, 244.49) mm, rotated rx 116.15 ry 10.69 rz 159.3 deg; joints [-82.754, -85.453, 5.12, 51.978, 67.463, 238.917, 323.242, 1043.223, 878.936]
  MoveL 247 to (-1905.15, -765.27, 245.28) mm, rotated rx 116.69 ry 11.84 rz 157.79 deg; joints [-80.801, -85.4, 5.12, 51.978, 67.685, 237.597, 307.925, 1064.218, 878.936]
  MoveL 248 to (-1920.07, -755.59, 245.8) mm, rotated rx 116.54 ry 13.96 rz 154.21 deg; joints [-76.669, -84.268, 5.12, 51.978, 68.333, 235.055, 294.651, 1087.678, 878.936]
  MoveL 249 to (-1936.55, -744.6, 246.59) mm, rotated rx 117.3 ry 14.46 rz 154.18 deg; joints [-76.319, -84.704, 5.115, 51.978, 68.33, 234.533, 279.92, 1105.811, 878.936]
  MoveL 250 to (-1953.29, -732.31, 247.11) mm, rotated rx 117.84 ry 16.33 rz 151.97 deg; joints [-73.456, -84.209, 5.115, 51.978, 68.735, 232.298, 265.773, 1131.121, 878.937]
  MoveL 251 to (-1970.03, -718.96, 247.63) mm, rotated rx 119.43 ry 18.55 rz 150.59 deg; joints [-70.944, -84.209, 5.115, 51.978, 68.922, 229.54, 253.758, 1160.86, 878.065]
  MoveL 252 to (-1985.47, -704.57, 248.42) mm, rotated rx 121.14 ry 21.67 rz 148.57 deg; joints [-67.504, -83.823, 5.115, 51.978, 69.435, 225.722, 243.533, 1193.696, 878.065]
  MoveL 253 to (-1999.33, -689.66, 248.94) mm, rotated rx 123.55 ry 25.55 rz 146.95 deg; joints [-63.932, -83.312, 5.115, 51.978, 70.018, 220.863, 235.374, 1227.247, 878.065]
  MoveL 254 to (-2011.37, -673.97, 249.2) mm, rotated rx 125.27 ry 28.99 rz 145.58 deg; joints [-60.974, -82.36, 5.115, 51.978, 70.638, 216.514, 225.531, 1253.692, 878.066]
  MoveL 255 to (-2021.83, -657.48, 249.73) mm, rotated rx 126.65 ry 32.81 rz 143.94 deg; joints [-58.014, -81.171, 5.115, 51.978, 71.714, 212.024, 214.928, 1279.919, 881.568]
  MoveL 256 to (-2030.73, -640.48, 249.99) mm, rotated rx 129.87 ry 38.4 rz 143.36 deg; joints [-55.173, -81.17, 5.115, 51.978, 74.019, 206.286, 210.6, 1320.448, 898.955]
  MoveL 257 to (-2038.31, -622.95, 250.25) mm, rotated rx 133.5 ry 41.83 rz 144.9 deg; joints [-54.014, -81.17, 5.115, 51.978, 74.826, 201.932, 205.757, 1348.927, 903.852]
  MoveL 258 to (-2044.86, -605.16, 250.51) mm, rotated rx 136.22 ry 44.73 rz 146.01 deg; joints [-53.117, -81.169, 5.115, 51.978, 75.904, 198.591, 200.748, 1376.032, 911.924]
  MoveL 259 to (-2050.35, -587.63, 250.77) mm, rotated rx 139.82 ry 47.8 rz 147.97 deg; joints [-52.368, -81.169, 5.115, 51.978, 76.973, 194.785, 196.535, 1402.504, 919.904]
  MoveL 260 to (-2055.06, -570.89, 250.77) mm, rotated rx 140.05 ry 48.32 rz 147.97 deg; joints [-52.233, -81.169, 5.115, 51.978, 77.328, 194.368, 191.837, 1420.94, 923.002]
  MoveL 261 to (-2059.24, -555.45, 250.51) mm, rotated rx 142.18 ry 50.48 rz 149.09 deg; joints [-51.799, -81.169, 5.115, 51.978, 78.403, 192.04, 187.953, 1442.515, 932.307]
  MoveL 262 to (-2063.17, -538.97, 250.25) mm, rotated rx 146.56 ry 52.95 rz 152.21 deg; joints [-51.473, -81.169, 5.115, 51.978, 79.183, 188.45, 184.455, 1465.105, 938.62]
  MoveL 263 to (-2067.09, -519.09, 249.99) mm, rotated rx 152.92 ry 55.88 rz 157.06 deg; joints [-51.208, -81.169, 5.115, 51.968, 80.218, 183.852, 180.543, 1492.039, 947.269]
  MoveL 264 to (-2070.49, -496.07, 248.68) mm, rotated rx 160.97 ry 58.61 rz 163.6 deg; joints [-51.133, -81.168, 5.115, 51.968, 81.326, 178.831, 176.419, 1521.73, 957.885]
  MoveL 265 to (-2073.11, -470.17, 246.33) mm, rotated rx 175.09 ry 61.1 rz 175.7 deg; joints [-51.133, -81.168, 5.115, 51.789, 82.481, 171.449, 172.9, 1554.477, 970.569]
  MoveL 266 to (-2074.42, -445.05, 241.62) mm, rotated rx -155.92 ry 61.09 rz -158.64 deg; joints [-51.133, -81.167, 5.115, 50.73, 84.306, 157.837, 170.546, 1584.998, 995.024]
  MoveL 267 to (-2074.68, -423.86, 234.81) mm, rotated rx -138.26 ry 55.89 rz -143.54 deg; joints [-51.133, -81.167, 5.063, 50.224, 84.017, 147.395, 170.546, 1610.096, 1002.289]
  MoveL 268 to (-2074.68, -405.55, 227.49) mm, rotated rx -140.14 ry 56.74 rz -145.08 deg; joints [-51.037, -80.262, 5.063, 50.224, 83.532, 148.048, 165.871, 1621.003, 1002.291]
  MoveL 269 to (-2074.68, -388.55, 221.47) mm, rotated rx -144.45 ry 57.99 rz -148.79 deg; joints [-50.748, -79.846, 5.063, 50.224, 83.079, 150.371, 164.925, 1633.847, 1002.292]
  MoveL 270 to (-2074.94, -372.33, 217.29) mm, rotated rx -159.01 ry 59.96 rz -161.63 deg; joints [-50.748, -79.846, 5.154, 51.131, 81.899, 157.799, 164.925, 1649.18, 992.867]
  MoveL 271 to (-2075.46, -355.58, 215.19) mm, rotated rx -177.04 ry 59.63 rz -177.44 deg; joints [-50.748, -79.846, 5.365, 51.866, 79.93, 166.353, 164.925, 1659.911, 976.121]
  MoveL 272 to (-2076.51, -337.27, 214.41) mm, rotated rx 173.1 ry 59.1 rz 174.07 deg; joints [-50.719, -79.846, 5.366, 51.866, 79.543, 171.386, 164.376, 1673.23, 973.417]
  MoveL 273 to (-2077.3, -315.82, 214.15) mm, rotated rx 170.18 ry 58.85 rz 171.57 deg; joints [-50.719, -79.846, 5.366, 51.856, 79.472, 172.916, 163.659, 1693.116, 973.147]
  MoveL 274 to (-2078.6, -291.75, 214.15) mm, rotated rx 172.21 ry 58.8 rz 173.32 deg; joints [-50.719, -80.06, 5.366, 51.865, 79.421, 172.045, 163.772, 1719.597, 973.147]
  MoveL 275 to (-2079.91, -264.8, 214.15) mm, rotated rx 172.81 ry 58.85 rz 173.84 deg; joints [-50.716, -80.06, 5.366, 51.865, 79.435, 171.729, 162.464, 1746.864, 973.258]
  MoveL 276 to (-2081.48, -234.72, 214.15) mm, rotated rx 170.75 ry 58.67 rz 172.08 deg; joints [-50.716, -80.06, 5.366, 51.853, 79.384, 172.814, 160.945, 1775.799, 972.881]
  MoveL 277 to (-2082.79, -201.75, 214.15) mm, rotated rx 173.18 ry 58.64 rz 174.17 deg; joints [-50.716, -80.269, 5.366, 51.871, 79.336, 171.721, 161.023, 1811.412, 972.88]
  MoveL 278 to (-2084.1, -165.91, 214.15) mm, rotated rx 171.88 ry 58.06 rz 173.09 deg; joints [-50.664, -80.269, 5.366, 51.871, 78.829, 172.461, 160.507, 1845.916, 968.254]
  MoveL 279 to (-2085.14, -127.19, 214.15) mm, rotated rx 171.61 ry 58.03 rz 172.86 deg; joints [-50.664, -80.269, 5.366, 51.868, 78.823, 172.608, 159.467, 1884.464, 968.216]
  MoveL 280 to (-2086.19, -85.86, 214.15) mm, rotated rx 173.05 ry 58.63 rz 174.06 deg; joints [-50.664, -80.268, 5.366, 51.818, 79.326, 171.795, 157.861, 1927.035, 972.886]
  MoveL 281 to (-2086.97, -43.48, 214.15) mm, rotated rx 177.72 ry 59.09 rz 178.04 deg; joints [-50.664, -80.268, 5.366, 51.813, 79.623, 169.357, 156.77, 1972.074, 975.54]
  MoveL 282 to (-2087.5, -0.05, 213.89) mm, rotated rx 177.84 ry 59.45 rz 178.14 deg; joints [-50.664, -80.268, 5.366, 51.746, 79.977, 169.297, 155.887, 2015.637, 979.19]
  MoveL 283 to (-2086.97, 43.38, 214.15) mm, rotated rx -178.76 ry 58.88 rz -178.94 deg; joints [-50.664, -80.937, 5.366, 51.795, 79.818, 168.065, 160.819, 2065.452, 979.19]
  MoveL 284 to (-2086.19, 86.02, 214.15) mm, rotated rx -174.38 ry 58.24 rz -175.22 deg; joints [-50.664, -81.481, 5.366, 51.89, 79.663, 166.155, 165.243, 2114.536, 979.189]
  MoveL 285 to (-2085.14, 127.1, 214.15) mm, rotated rx -171.85 ry 58.06 rz -173.07 deg; joints [-50.664, -81.521, 5.366, 51.935, 79.651, 164.832, 166.568, 2157.45, 979.189]
  MoveL 286 to (-2084.1, 166.08, 214.15) mm, rotated rx -173.39 ry 58.18 rz -174.38 deg; joints [-50.665, -81.476, 5.526, 51.934, 79.547, 165.494, 166.568, 2194.248, 979.189]
  MoveL 287 to (-2082.79, 201.92, 214.15) mm, rotated rx -173.76 ry 58.68 rz -174.66 deg; joints [-50.665, -81.148, 5.526, 51.853, 79.808, 165.494, 165.499, 2227.308, 980.805]
  MoveL 288 to (-2081.48, 234.62, 214.15) mm, rotated rx -172.81 ry 58.85 rz -173.84 deg; joints [-50.665, -80.956, 5.526, 51.832, 79.904, 164.877, 165.49, 2259.051, 981.212]
  MoveL 289 to (-2079.91, 264.7, 214.15) mm, rotated rx -172.21 ry 58.8 rz -173.32 deg; joints [-50.665, -80.968, 5.526, 51.839, 79.899, 164.57, 167.148, 2289.559, 981.212]
  MoveL 290 to (-2078.6, 291.65, 214.15) mm, rotated rx -173.07 ry 58.87 rz -174.06 deg; joints [-50.665, -80.92, 5.743, 51.864, 79.753, 164.813, 167.148, 2314.457, 981.212]
  MoveL 291 to (-2077.3, 315.98, 214.15) mm, rotated rx -167.48 ry 58.53 rz -169.28 deg; joints [-50.627, -80.8, 5.743, 51.864, 79.764, 161.797, 167.867, 2340.716, 981.212]
  MoveL 292 to (-2076.51, 337.17, 214.41) mm, rotated rx -176.78 ry 59.33 rz -177.23 deg; joints [-50.627, -80.592, 5.877, 51.784, 79.764, 166.402, 166.611, 2354.73, 981.212]
  MoveL 293 to (-2075.46, 355.75, 215.19) mm, rotated rx -179.41 ry 59.59 rz -179.49 deg; joints [-50.627, -80.422, 6.045, 51.77, 79.764, 167.488, 165.7, 2369.851, 981.212]
  MoveL 294 to (-2074.94, 372.49, 217.29) mm, rotated rx 159.35 ry 60.05 rz 161.92 deg; joints [-50.602, -78.955, 6.045, 51.77, 80.913, 176.792, 156.254, 2369.851, 986.821]
  MoveL 295 to (-2074.68, 388.71, 221.47) mm, rotated rx 145.03 ry 58.19 rz 149.27 deg; joints [-50.034, -77.66, 6.771, 51.77, 80.913, 182.687, 147.227, 2370.378, 986.821]
  MoveL 296 to (-2074.68, 405.45, 227.49) mm, rotated rx 139.35 ry 56.43 rz 144.42 deg; joints [-49.786, -77.66, 6.997, 51.77, 80.913, 186.044, 147.117, 2384.527, 983.579]
  MoveL 297 to (-2074.68, 423.77, 234.81) mm, rotated rx 137.92 ry 55.72 rz 143.28 deg; joints [-49.786, -77.66, 7.006, 51.818, 80.788, 187.093, 147.117, 2402.059, 975.405]
  MoveL 298 to (-2074.42, 444.96, 241.62) mm, rotated rx 151.83 ry 60.26 rz 155.07 deg; joints [-49.786, -77.66, 7.054, 51.34, 80.882, 178.512, 147.118, 2426.09, 968.69]
  MoveL 299 to (-2073.11, 470.33, 246.33) mm, rotated rx 177.22 ry 61.46 rz 177.55 deg; joints [-50.064, -77.66, 7.054, 51.34, 79.143, 166.296, 148.131, 2456.089, 946.722]
  MoveL 300 to (-2070.49, 495.97, 248.68) mm, rotated rx -167.94 ry 59.94 rz -169.53 deg; joints [-50.064, -78.796, 7.054, 51.34, 78.86, 159.833, 158.235, 2495.402, 944.359]
  MoveL 301 to (-2067.09, 518.99, 249.99) mm, rotated rx -158.27 ry 57.84 rz -161.35 deg; joints [-50.063, -79.749, 7.054, 51.486, 78.731, 155.173, 167.896, 2530.739, 944.357]
  MoveL 302 to (-2063.17, 539.14, 250.25) mm, rotated rx -150.74 ry 54.88 rz -155.38 deg; joints [-50.063, -80.985, 7.054, 51.936, 78.422, 151.074, 180.225, 2567.125, 944.357]
  MoveL 303 to (-2059.24, 555.62, 250.51) mm, rotated rx -145.72 ry 51.95 rz -151.78 deg; joints [-50.063, -82.241, 7.054, 52.57, 78.097, 147.936, 192.927, 2600.767, 944.357]
  MoveL 304 to (-2055.06, 571.05, 250.77) mm, rotated rx -142.72 ry 49.84 rz -149.82 deg; joints [-50.063, -83.089, 7.054, 53.115, 77.867, 145.808, 203.233, 2628.798, 944.357]
  MoveL 305 to (-2050.35, 587.54, 250.77) mm, rotated rx -140.65 ry 48.41 rz -148.48 deg; joints [-50.063, -83.51, 7.054, 53.497, 77.724, 144.162, 211.151, 2652.932, 944.357]
  MoveL 306 to (-2044.86, 605.06, 250.51) mm, rotated rx -139.2 ry 47.33 rz -147.6 deg; joints [-50.063, -83.789, 7.054, 53.813, 77.599, 142.924, 218.896, 2676.131, 944.357]
  MoveL 307 to (-2038.31, 622.85, 250.25) mm, rotated rx -135.6 ry 44.51 rz -145.53 deg; joints [-50.063, -84.425, 7.054, 54.678, 77.33, 139.619, 230.812, 2708.498, 944.357]
  MoveL 308 to (-2030.73, 640.64, 249.99) mm, rotated rx -132.64 ry 42.22 rz -143.88 deg; joints [-50.063, -84.699, 7.054, 55.394, 77.167, 136.612, 241.278, 2736.646, 944.357]
  MoveL 309 to (-2021.83, 657.65, 249.73) mm, rotated rx -129.72 ry 37.19 rz -143.96 deg; joints [-50.063, -86.724, 7.054, 57.951, 76.411, 132.949, 268.323, 2792.935, 944.357]
  MoveL 310 to (-2011.37, 673.87, 249.2) mm, rotated rx -127.3 ry 32.91 rz -144.5 deg; joints [-50.063, -88.114, 7.054, 60.551, 75.761, 129.455, 294.111, 2843.709, 944.357]
  MoveL 311 to (-1999.33, 689.57, 248.94) mm, rotated rx -124.69 ry 28.89 rz -145.09 deg; joints [-50.063, -88.971, 7.054, 63.274, 75.305, 125.495, 319.241, 2891.101, 944.356]
  MoveL 312 to (-1985.47, 704.74, 248.42) mm, rotated rx -121.89 ry 24.43 rz -146.38 deg; joints [-50.063, -89.657, 7.054, 66.851, 74.887, 120.804, 349.02, 2943.712, 944.356]
  MoveL 313 to (-1970.03, 718.87, 247.63) mm, rotated rx -119.82 ry 20.17 rz -148.97 deg; joints [-50.063, -90.454, 7.054, 71.218, 74.38, 116.727, 386.328, 3000.967, 944.356]
  MoveL 314 to (-1953.29, 732.47, 247.11) mm, rotated rx -118.13 ry 17.95 rz -150.04 deg; joints [-49.142, -90.454, 7.054, 72.595, 74.38, 113.866, 417.395, 3030.172, 945.554]
  MoveL 315 to (-1936.55, 744.77, 246.59) mm, rotated rx -117.53 ry 15.62 rz -152.67 deg; joints [-49.142, -91.119, 7.054, 75.884, 73.947, 112.142, 454.142, 3072.913, 945.554]
  MoveL 316 to (-1920.07, 755.75, 245.8) mm, rotated rx -117.03 ry 13.91 rz -154.78 deg; joints [-49.142, -91.505, 7.054, 78.52, 73.639, 110.738, 486.693, 3106.564, 945.554]
  MoveL 317 to (-1905.15, 765.17, 245.28) mm, rotated rx -117.24 ry 13.48 rz -155.65 deg; joints [-49.142, -91.756, 7.054, 79.367, 73.35, 110.738, 508.186, 3123.487, 944.998]
  MoveL 318 to (-1888.15, 774.33, 244.49) mm, rotated rx -116.28 ry 11.39 rz -158.19 deg; joints [-49.142, -91.932, 7.052, 82.749, 73.202, 108.536, 544.925, 3158.717, 944.997]
  MoveL 319 to (-1866.7, 785.05, 243.45) mm, rotated rx -115.72 ry 10.66 rz -158.98 deg; joints [-47.982, -91.932, 7.052, 82.749, 73.217, 107.588, 579.221, 3172.396, 946.904]
  MoveL 320 to (-1838.96, 796.83, 242.4) mm, rotated rx -114.64 ry 9.12 rz -160.94 deg; joints [-45.614, -91.932, 7.052, 83.065, 73.217, 105.632, 635.311, 3191.378, 949.218]
  MoveL 321 to (-1802.6, 810.17, 240.83) mm, rotated rx -112.4 ry 7.73 rz -161.94 deg; joints [-44.518, -91.932, 7.052, 83.862, 74.329, 103.158, 687.201, 3214.976, 962.097]
  MoveL 322 to (-1760.74, 824.04, 239.26) mm, rotated rx -111.15 ry 6.42 rz -163.88 deg; joints [-41.972, -91.932, 7.052, 83.862, 74.638, 101.326, 757.8, 3232.855, 967.926]
  MoveL 323 to (-1716.01, 837.12, 237.69) mm, rotated rx -109.45 ry 5.35 rz -165.22 deg; joints [-40.071, -91.932, 7.052, 83.862, 75.475, 99.464, 823.368, 3249.613, 978.592]
  MoveL 324 to (-1669.7, 849.93, 236.12) mm, rotated rx -107.53 ry 4.62 rz -165.7 deg; joints [-39.158, -91.932, 7.052, 83.863, 76.705, 97.807, 878.928, 3265.927, 992.719]
  Set speed (1000.0 mm/s)
  MoveL 325 to (-1669.7, 849.93, 236.12) mm, rotated rx -107.53 ry 4.62 rz -165.7 deg; joints [-39.158, -91.932, 7.052, 83.863, 76.705, 97.807, 878.928, 3265.927, 992.719]
  MoveL 326 to (-1695.61, 941.74, 266.15) mm, rotated rx -107.53 ry 4.62 rz -165.7 deg; joints [-39.158, -91.932, 7.052, 83.863, 76.705, 97.807, 853.022, 3357.728, 962.694]

--- program Trunk_C (robot ABB IRB 1300-10/1.15) ---
  Smooth(1)
  Set speed (1000.0 mm/s)
  Set Ref.: Trunk
  Set Tool: Generic Paint Sprayer
  Show Generic Paint Sprayer
  MoveJ 1 to (5.82, -17.96, 97.39) mm, rotated rx 3.37 ry -10.35 rz -90.2 deg; joints [-81.249, 102.668, -200.517, 127.068, 82.563, -85.716, 20.249, 2120.861, 930.715]
  MoveL 2 to (5.82, -17.96, 97.39) mm, rotated rx 3.37 ry -10.35 rz -90.2 deg; joints [-81.249, 102.661, -200.517, 127.066, 82.558, -85.71, 20.249, 2120.898, 930.657]
  MoveL 3 to (0, 0, 195.59) mm, rotated rx 3.37 ry -10.35 rz -90.2 deg; joints [-81.249, 102.661, -200.517, 127.066, 82.558, -85.71, 116.053, 2092.818, 936.418]
  MoveL 4 to (0, 0, 195.59) mm, rotated rx 3.37 ry -10.35 rz -90.2 deg; joints [-81.249, 102.661, -200.517, 127.066, 82.558, -85.71, 116.053, 2092.818, 936.418]
  Set speed (200.0 mm/s)
  MoveL 5 to (0, 100, 183.28) mm, rotated rx 4.4 ry -4.25 rz -90.13 deg; joints [-86.651, 102.661, -200.644, 126.277, 81.606, -86.022, 116.053, 1943.952, 926.891]
  MoveL 6 to (0, 200, 178.84) mm, rotated rx 3.06 ry -1.77 rz -90.1 deg; joints [-89.2, 101.304, -200.644, 126.277, 81.918, -84.247, 114.795, 1831.463, 926.891]
  MoveL 7 to (0, 300, 178.89) mm, rotated rx 3.77 ry 1.04 rz -90.08 deg; joints [-91.442, 101.304, -200.74, 125.636, 81.314, -84.45, 114.795, 1710.076, 920.567]
  MoveL 8 to (0, 400, 182.92) mm, rotated rx 3.05 ry 3.15 rz -90.04 deg; joints [-92.986, 101.304, -200.734, 125.13, 81.975, -84.015, 114.795, 1593.285, 926.079]
  MoveL 9 to (0, 500, 189.58) mm, rotated rx 3.08 ry 4.3 rz -90.02 deg; joints [-93.81, 101.304, -200.734, 124.801, 81.99, -83.984, 114.795, 1483.964, 925.485]
  MoveL 10 to (0, 600, 197.8) mm, rotated rx 2.6 ry 7.21 rz -90 deg; joints [-95.162, 100.893, -200.734, 123.236, 82.372, -83.249, 114.795, 1361.904, 925.866]
  MoveL 11 to (0, 700, 210.65) mm, rotated rx 3.09 ry 7.59 rz -90.03 deg; joints [-95.162, 100.893, -201.006, 122.78, 81.864, -83.249, 115.815, 1259.807, 921.904]
  MoveL 12 to (0, 800, 225.02) mm, rotated rx 3.08 ry 8.74 rz -90.06 deg; joints [-95.187, 100.893, -201.006, 121.66, 82.047, -83.161, 115.815, 1148.837, 921.711]
  MoveL 13 to (0, 900, 242.24) mm, rotated rx 3.81 ry 10.85 rz -90.09 deg; joints [-95.2, 100.893, -201.227, 119.471, 81.63, -83.161, 115.815, 1030.666, 915.578]
  MoveL 14 to (0, 1000, 263.68) mm, rotated rx 5.07 ry 13.41 rz -90.12 deg; joints [-95.2, 100.893, -201.706, 116.723, 80.732, -83.161, 119.571, 909.641, 905.365]
  MoveL 15 to (0, 1100, 290) mm, rotated rx 6.24 ry 16.08 rz -89.82 deg; joints [-95.2, 100.893, -201.767, 113.895, 80.071, -83.161, 129.337, 783.636, 894.572]
  Set speed (1000.0 mm/s)
  MoveL 16 to (0, 1100, 290) mm, rotated rx 6.24 ry 16.08 rz -89.82 deg; joints [-95.2, 100.893, -201.767, 113.895, 80.071, -83.161, 129.337, 783.636, 894.572]
  MoveL 17 to (10.79, 1127.56, 194.48) mm, rotated rx 6.24 ry 16.08 rz -89.82 deg; joints [-95.2, 100.893, -201.767, 113.895, 80.071, -83.161, 31.476, 766.175, 883.702]
  Set speed (1000.0 mm/s)
  MoveL 18 to (67.64, 1129.95, 194.57) mm, rotated rx -4.11 ry 17.5 rz -89.62 deg; joints [-95.2, 100.893, -201.767, 113.96, 89.111, -77.809, 26.478, 750.723, 915.458]
  MoveL 19 to (75, 1100, 289.7) mm, rotated rx -4.11 ry 17.5 rz -89.62 deg; joints [-95.2, 100.893, -201.767, 113.96, 89.111, -77.809, 124.201, 770.659, 908.189]
  MoveL 20 to (75, 1100, 289.7) mm, rotated rx -4.11 ry 17.5 rz -89.62 deg; joints [-95.2, 100.893, -201.767, 113.96, 89.111, -77.809, 124.201, 770.659, 908.189]
  Set speed (200.0 mm/s)
  MoveL 21 to (75, 1000, 262.1) mm, rotated rx -5.7 ry 14.12 rz -89.62 deg; joints [-95.2, 100.893, -201.188, 117.583, 90.137, -77.809, 116.908, 899.97, 920.835]
  MoveL 22 to (75, 900, 239.63) mm, rotated rx -4.57 ry 11.49 rz -87.14 deg; joints [-95.2, 102.696, -201.188, 120.034, 88.858, -77.81, 112.727, 1017.527, 920.314]
  MoveL 23 to (75, 800, 221.68) mm, rotated rx -5.34 ry 9.29 rz -87.12 deg; joints [-95.153, 102.695, -200.958, 122.292, 89.252, -77.81, 112.727, 1136.937, 925.754]
  MoveL 24 to (75, 700, 206.84) mm, rotated rx -5.72 ry 8.19 rz -86.8 deg; joints [-95.138, 102.695, -200.5, 123.436, 89.532, -77.81, 112.727, 1244.6, 927.254]
  MoveL 25 to (75, 600, 193.75) mm, rotated rx -6.16 ry 7.55 rz -87.06 deg; joints [-95.13, 102.604, -200.5, 124.136, 89.846, -77.81, 112.727, 1351.468, 930.969]
  MoveL 26 to (75, 500, 185.55) mm, rotated rx -5.85 ry 4.6 rz -85.52 deg; joints [-93.809, 103.701, -200.32, 125.699, 89.347, -77.81, 112.727, 1470.008, 930.969]
  MoveL 27 to (75, 400, 179.15) mm, rotated rx -5.99 ry 3.32 rz -85.57 deg; joints [-92.92, 103.665, -200.32, 126.102, 89.347, -77.822, 112.727, 1580.554, 931.542]
  MoveL 28 to (75, 300, 175.65) mm, rotated rx -5.11 ry 1.19 rz -84.9 deg; joints [-91.451, 105.01, -200.32, 126.598, 88.879, -78.872, 112.727, 1690.665, 931.541]
  MoveL 29 to (75, 200, 176.25) mm, rotated rx -5.59 ry -1.42 rz -84.92 deg; joints [-89.251, 105.01, -200.213, 127.065, 89.138, -78.866, 112.727, 1810.509, 933.966]
  MoveL 30 to (75, 100, 181.63) mm, rotated rx -4.89 ry -3.78 rz -84.22 deg; joints [-87.026, 106.265, -200.213, 127.065, 88.731, -79.754, 115.435, 1922.634, 933.963]
  MoveL 31 to (75, 0, 195.43) mm, rotated rx -3.81 ry -11.34 rz -83.77 deg; joints [-81.006, 108.305, -200.213, 128.425, 88.107, -82.066, 115.435, 2073.703, 933.933]
  Set speed (1000.0 mm/s)
  MoveL 32 to (75, 0, 195.43) mm, rotated rx -3.81 ry -11.34 rz -83.77 deg; joints [-81.006, 108.305, -200.213, 128.425, 88.107, -82.066, 115.435, 2073.703, 933.933]
  MoveL 33 to (70.53, -20.22, 97.6) mm, rotated rx -3.81 ry -11.34 rz -83.77 deg; joints [-81.006, 108.305, -200.213, 128.425, 88.107, -82.066, 20.229, 2103.954, 938.472]
  Set speed (1000.0 mm/s)
  MoveL 34 to (224.3, -61.4, 171.25) mm, rotated rx -68.37 ry -43.71 rz 35.1 deg; joints [-39.191, 151.79, -172.14, 171.412, 88.107, -89.491, 21.941, 2103.953, 850.723]
  MoveL 35 to (150, 0, 197.9) mm, rotated rx -68.37 ry -43.71 rz 35.1 deg; joints [-39.191, 151.79, -172.14, 171.412, 88.107, -89.491, 42.046, 2039.88, 924.82]
  MoveL 36 to (150, 0, 197.9) mm, rotated rx -68.37 ry -43.71 rz 35.1 deg; joints [-39.191, 151.79, -172.14, 171.412, 88.107, -89.491, 42.046, 2039.88, 924.82]
  Set speed (200.0 mm/s)
  MoveL 37 to (150, 100, 176.5) mm, rotated rx -6.65 ry -1.9 rz -31.75 deg; joints [-82.988, 150.879, -195.912, 121.767, 88.107, -75.985, 42.044, 1775.32, 1100]
  MoveL 38 to (150, 200, 168.83) mm, rotated rx -2.6 ry 3.06 rz -31.84 deg; joints [-86.723, 149.043, -195.912, 118.606, 87.146, -74.604, 42.044, 1618.084, 1100]
  MoveL 39 to (150, 300, 169.73) mm, rotated rx -0.66 ry 3.24 rz -31.84 deg; joints [-87.706, 149.046, -195.912, 118.696, 86.165, -75.212, 42.043, 1503.214, 1092.233]
  MoveL 40 to (150, 400, 172.48) mm, rotated rx -0.15 ry 4.49 rz -31.74 deg; joints [-88.533, 149.046, -195.912, 117.946, 86.507, -75.013, 39.348, 1393.761, 1098.767]
  MoveL 41 to (150, 500, 178.13) mm, rotated rx 1.19 ry 5.7 rz -31.7 deg; joints [-89.35, 149.046, -196.245, 117.032, 86.03, -75.013, 39.348, 1280.386, 1099.936]
  Set speed (1000.0 mm/s)
  MoveL 42 to (150, 500, 178.13) mm, rotated rx 1.19 ry 5.7 rz -31.7 deg; joints [-89.35, 149.046, -196.245, 117.032, 86.03, -75.013, 39.348, 1280.386, 1099.936]
  MoveL 43 to (142.64, 506.98, 78.64) mm, rotated rx 1.19 ry 5.7 rz -31.66 deg; joints [-94.245, 148.306, -196.245, 120.534, 88.546, -72.733, 0, 1283.545, 1100]
  Set speed (1000.0 mm/s)
  MoveL 44 to (143.25, 714.01, 100.59) mm, rotated rx 4.83 ry 7.54 rz -31.48 deg; joints [-94.825, 148.306, -196.245, 118.28, 86.372, -74.165, 0.001, 1040.894, 1095.98]
  MoveL 45 to (150, 700, 199.37) mm, rotated rx 4.83 ry 7.54 rz -31.48 deg; joints [-94.825, 148.306, -196.245, 118.28, 86.372, -74.165, 99.707, 1044.588, 1089.267]
  MoveL 46 to (150, 700, 199.37) mm, rotated rx 4.87 ry 7.51 rz -31.14 deg; joints [-94.826, 148.381, -196.245, 118.238, 86.243, -73.93, 99.707, 1043.629, 1089.279]
  Set speed (200.0 mm/s)
  MoveL 47 to (150, 800, 214.95) mm, rotated rx 6.43 ry 7.71 rz -31.11 deg; joints [-94.871, 148.381, -196.245, 117.713, 85.032, -74.646, 104.839, 930.339, 1083.42]
  MoveL 48 to (150, 900, 233.48) mm, rotated rx 7.85 ry 8.45 rz -30.95 deg; joints [-94.871, 148.381, -196.246, 116.656, 84.025, -75.181, 110.911, 814.917, 1082.239]
  MoveL 49 to (150, 1000, 254.37) mm, rotated rx 9.73 ry 11.24 rz -30.42 deg; joints [-94.871, 148.381, -196.75, 113.429, 82.997, -75.181, 113.765, 688.961, 1092.754]
  MoveL 50 to (150, 1100, 285.02) mm, rotated rx 15.79 ry 11.38 rz -30.24 deg; joints [-94.925, 148.407, -196.75, 112.05, 77.934, -77.853, 140.904, 541.747, 1066.066]
  Set speed (1000.0 mm/s)
  MoveL 51 to (150, 1100, 285.02) mm, rotated rx 15.79 ry 11.38 rz -30.24 deg; joints [-94.925, 148.407, -196.75, 112.05, 77.934, -77.853, 140.904, 541.747, 1066.066]
  MoveL 52 to (147.3, 1133.07, 190.69) mm, rotated rx 15.79 ry 11.38 rz -30.24 deg; joints [-94.925, 148.407, -196.75, 112.05, 77.934, -77.853, 43.644, 518.641, 1068.659]
  Set speed (1000.0 mm/s)
  MoveL 53 to (229.18, 919.28, 136.73) mm, rotated rx 10.7 ry 3.91 rz -32.08 deg; joints [-94.925, 148.407, -195.888, 120.751, 80.838, -77.852, 31.544, 806.698, 958.042]
  MoveL 54 to (225, 900, 234.76) mm, rotated rx 10.7 ry 3.91 rz -32.08 deg; joints [-94.925, 148.407, -195.888, 120.751, 80.838, -77.852, 131.049, 815.682, 962.282]
  MoveL 55 to (225, 900, 234.76) mm, rotated rx 8.72 ry 7.34 rz -52.03 deg; joints [-94.925, 142.985, -195.888, 121.299, 88.033, -90.753, 124.527, 862.143, 962.282]
  Set speed (200.0 mm/s)
  MoveL 56 to (225, 800, 217.13) mm, rotated rx 9.67 ry 3.88 rz -52.44 deg; joints [-94.369, 142.985, -195.888, 124.365, 86.884, -91.456, 124.527, 982.115, 938.152]
  MoveL 57 to (225, 700, 202.35) mm, rotated rx 8.96 ry 2.98 rz -52.58 deg; joints [-94.369, 142.971, -195.888, 125.266, 87.503, -91.121, 123.402, 1093.142, 938.693]
  MoveL 58 to (225, 600, 189.34) mm, rotated rx 8.85 ry 2.39 rz -52.39 deg; joints [-94.369, 142.971, -195.56, 125.829, 87.665, -91.121, 123.345, 1195.648, 937.556]
  MoveL 59 to (225, 500, 181.24) mm, rotated rx 4.92 ry 1.35 rz -52.47 deg; joints [-93.975, 142.964, -195.56, 126.545, 90.85, -89.263, 123.344, 1323.083, 959.284]
  MoveL 60 to (225, 400, 174.94) mm, rotated rx 3.6 ry 0.9 rz -52.44 deg; joints [-93.497, 142.964, -195.56, 126.629, 91.72, -88.714, 123.334, 1432.531, 966.157]
  MoveL 61 to (225, 300, 171.21) mm, rotated rx 1.64 ry 0.76 rz -52.45 deg; joints [-92.891, 142.954, -195.56, 126.332, 93.11, -87.934, 123.334, 1543.106, 979.029]
  Set speed (1000.0 mm/s)
  MoveL 62 to (225, 300, 171.21) mm, rotated rx 1.64 ry 0.76 rz -52.45 deg; joints [-92.891, 142.954, -195.56, 126.332, 93.11, -87.934, 123.334, 1543.106, 979.029]
  MoveL 63 to (226.47, 302.79, 71.26) mm, rotated rx 1.81 ry 0.05 rz -29.31 deg; joints [-95.547, 149.146, -195.56, 126.333, 86.829, -71.804, 51.369, 1498.461, 979.029]
  Set speed (1000.0 mm/s)
  MoveL 64 to (367.99, -36.42, 198.34) mm, rotated rx 3.76 ry -50.37 rz -33.06 deg; joints [-81.345, 131.225, -165.038, 169.074, 85.783, -93.995, 375.631, 1750.09, 538.837]
  MoveL 65 to (300, 0, 261.98) mm, rotated rx 3.76 ry -50.37 rz -33.06 deg; joints [-81.345, 131.225, -165.038, 169.074, 85.783, -93.995, 435.125, 1707.035, 606.709]
  MoveL 66 to (300, 0, 261.98) mm, rotated rx 3.76 ry -50.37 rz -33.06 deg; joints [-81.345, 131.225, -165.038, 169.074, 85.783, -93.995, 435.125, 1707.035, 606.709]
  Set speed (200.0 mm/s)
  MoveL 67 to (300, 100, 226.55) mm, rotated rx 20.15 ry -38.1 rz -41.72 deg; joints [-90.05, 131.49, -165.038, 162.967, 82.074, -98.516, 435.125, 1534.268, 606.709]
  MoveL 68 to (300, 200, 215.25) mm, rotated rx 23.07 ry -34.87 rz -40.11 deg; joints [-92.829, 131.95, -165.037, 161.147, 79.408, -97.864, 435.124, 1397.375, 606.708]
  MoveL 69 to (300, 300, 213.38) mm, rotated rx 26.4 ry -32.38 rz -41.29 deg; joints [-94.303, 132.067, -165.038, 160.072, 78.314, -99.409, 435.124, 1279.404, 606.708]
  MoveL 70 to (300, 400, 216.67) mm, rotated rx 26.48 ry -31.14 rz -40.56 deg; joints [-95.378, 132.067, -165.037, 159.146, 78.012, -98.497, 435.124, 1171.901, 608.809]
  MoveL 71 to (300, 500, 222.55) mm, rotated rx 27.02 ry -30.26 rz -40.88 deg; joints [-95.979, 131.982, -165.038, 158.7, 78.008, -98.589, 435.124, 1069.197, 609.084]
  MoveL 72 to (300, 600, 230.2) mm, rotated rx 28.84 ry -28.9 rz -40.06 deg; joints [-96.528, 132.217, -165.038, 157.666, 76.259, -99.079, 435.124, 947.253, 609.084]
  MoveL 73 to (300, 700, 243.15) mm, rotated rx 29.51 ry -28.63 rz -40.55 deg; joints [-96.528, 132.285, -165.038, 157.666, 76.199, -99.761, 437.984, 845.015, 609.084]
  MoveL 74 to (300, 800, 257.52) mm, rotated rx 30.64 ry -28.81 rz -40.68 deg; joints [-96.528, 132.626, -165.038, 158.083, 75.642, -100.529, 446.684, 737.939, 609.084]
  MoveL 75 to (300, 900, 275.04) mm, rotated rx 33.53 ry -27.5 rz -42.8 deg; joints [-96.528, 132.83, -165.038, 158.095, 75.328, -103.523, 455.566, 630.54, 609.084]
  MoveL 76 to (300, 1000, 298.86) mm, rotated rx 35.17 ry -24.77 rz -40.68 deg; joints [-96.627, 132.83, -165.038, 155.311, 72.387, -103.923, 455.566, 493.244, 611.181]
  MoveL 77 to (300, 1100, 335.43) mm, rotated rx 40.69 ry -23.26 rz -39.34 deg; joints [-96.627, 133.603, -165.038, 154.938, 67.49, -107.1, 492.895, 338.537, 611.181]
  Set speed (1000.0 mm/s)
  MoveL 78 to (300, 1100, 335.43) mm, rotated rx 40.69 ry -23.26 rz -39.34 deg; joints [-96.627, 133.603, -165.038, 154.938, 67.49, -107.1, 492.895, 338.537, 611.181]
  MoveL 79 to (364.49, 1131.44, 265.77) mm, rotated rx 40.69 ry -23.26 rz -39.34 deg; joints [-96.627, 133.718, -165.153, 154.938, 67.49, -107.1, 420.274, 315.502, 547.432]

--- program Trunk_Top_C (robot ABB IRB 1300-10/1.15) ---
  Smooth(1)
  Set speed (1000.0 mm/s)
  Set Ref.: Trunk
  Set Tool: Generic Paint Sprayer
  Show Generic Paint Sprayer
  MoveJ 1 to (1053.45, 1050.9, 272.58) mm, rotated rx 42.19 ry -24.4 rz -21.91 deg; joints [-68.905, 132.2, -165.153, 105.882, 75.627, 78.443, 47.258, 1676.865, 605.202]
  MoveL 2 to (1053.45, 1050.9, 272.58) mm, rotated rx 42.19 ry -24.4 rz -21.91 deg; joints [-68.905, 132.2, -165.153, 105.882, 75.627, 78.443, 47.258, 1676.865, 605.202]
  MoveL 3 to (1000, 1000, 340.05) mm, rotated rx -24.01 ry -42.38 rz 77.06 deg; joints [0, 69.901, -170.076, 54.11, 82.773, 207.011, 9.386, 2714.379, 0.001]
  MoveL 4 to (1000, 1000, 340.05) mm, rotated rx -24.01 ry -42.38 rz 77.06 deg; joints [0, 69.901, -170.076, 54.11, 82.773, 207.011, 9.386, 2714.379, 0.001]
  Set speed (200.0 mm/s)
  MoveL 5 to (1000, 900, 183.05) mm, rotated rx -5.71 ry -7.49 rz 90.27 deg; joints [14.805, 112.588, -172.639, 106.526, 36.703, 140.958, 0, 2714.377, 0]
  MoveL 6 to (1000, 800, 174.67) mm, rotated rx -6.59 ry -3.49 rz 90.12 deg; joints [18.243, 114.854, -172.639, 111.489, 32.385, 133.587, 0, 2633.3, 0]
  MoveL 7 to (1000, 700, 170.36) mm, rotated rx -6.5 ry -1.9 rz 90.06 deg; joints [18.665, 115.879, -172.639, 115.194, 31.625, 129.661, 0, 2526.902, 0]
  MoveL 8 to (1000, 600, 167.93) mm, rotated rx -6.44 ry -0.83 rz 90.05 deg; joints [18.86, 116.546, -172.639, 117.816, 31.258, 127.01, 0, 2421.234, 0]
  MoveL 9 to (1000, 500, 167.2) mm, rotated rx -6.45 ry 0.4 rz 90.04 deg; joints [19.314, 117.106, -172.639, 120.448, 30.636, 124.237, 0.885, 2317.72, 0]
  MoveL 10 to (1000, 400, 168.48) mm, rotated rx -6.45 ry 1.1 rz 90.09 deg; joints [19.719, 117.328, -172.639, 121.851, 30.227, 122.694, 2.712, 2217.7, 0.004]
  MoveL 11 to (1000, 300, 171.79) mm, rotated rx -6.43 ry 2.32 rz 90.06 deg; joints [20.449, 117.542, -172.639, 124.13, 29.421, 120.08, 6.176, 2117.645, 0.003]
  MoveL 12 to (1000, 200, 176.79) mm, rotated rx -6.5 ry 3.39 rz 90.06 deg; joints [21.362, 117.549, -172.639, 125.853, 28.486, 117.908, 10.561, 2021.276, 0.002]
  MoveL 13 to (1000, 100, 183.69) mm, rotated rx -6.57 ry 5 rz 90.15 deg; joints [22.813, 117.529, -172.612, 128.747, 27.187, 114.328, 18.384, 1927.653, 0.002]
  MoveL 14 to (1000, 0, 194.67) mm, rotated rx -5.71 ry 8.97 rz 89.75 deg; joints [24.407, 117.78, -172.612, 138.055, 26.133, 104.049, 33.858, 1814.006, 0]
  Set speed (1000.0 mm/s)
  MoveL 15 to (1000, 0, 194.67) mm, rotated rx -5.71 ry 8.97 rz 89.75 deg; joints [24.407, 117.78, -172.612, 138.055, 26.133, 104.049, 33.858, 1814.006, 0]
  MoveL 16 to (1009.89, -15.56, 96.38) mm, rotated rx -5.71 ry 8.97 rz 89.75 deg; joints [25.361, 126.017, -172.463, 147.269, 32.463, 92.662, 20.877, 1816.347, 6.741]
  Set speed (1000.0 mm/s)
  MoveL 17 to (913.66, -14.01, 83.62) mm, rotated rx -7.87 ry 8.11 rz 89.83 deg; joints [24.704, 126.871, -172.725, 145.766, 31.383, 95.44, 95.907, 1816.347, 6.742]
  MoveL 18 to (900, 0, 181.69) mm, rotated rx -7.87 ry 8.11 rz 89.83 deg; joints [24.695, 126.86, -172.718, 145.761, 31.383, 95.454, 111.319, 1828.983, 104.598]
  MoveL 19 to (900, 0, 181.69) mm, rotated rx -7.87 ry 8.11 rz 89.83 deg; joints [24.695, 126.86, -172.718, 145.761, 31.383, 95.454, 111.319, 1828.983, 104.598]
  Set speed (200.0 mm/s)
  MoveL 20 to (900, 100, 170.1) mm, rotated rx -8.23 ry 5.17 rz 89.96 deg; joints [21.85, 126.989, -172.898, 139.621, 32.562, 103.18, 92.356, 1915.011, 104.597]
  MoveL 21 to (900, 200, 162.09) mm, rotated rx -8.64 ry 3.98 rz 91.28 deg; joints [21.489, 127.239, -173.105, 137.261, 33.224, 106.701, 92.356, 2021.553, 104.597]
  MoveL 22 to (900, 300, 156.71) mm, rotated rx -8.83 ry 2.75 rz 91.3 deg; joints [20.388, 127.193, -173.105, 134.925, 33.866, 109.578, 85.022, 2116.694, 104.598]
  MoveL 23 to (900, 400, 153.25) mm, rotated rx -8.72 ry 1.4 rz 92.07 deg; joints [19.592, 127.025, -173.105, 132.596, 35.003, 112.7, 85.022, 2217.803, 105.16]
  MoveL 24 to (900, 500, 151.96) mm, rotated rx -8.74 ry 0.71 rz 91.99 deg; joints [18.776, 126.972, -173.105, 131.447, 35.548, 114.206, 80.599, 2311.833, 107.239]
  MoveL 25 to (900, 600, 152.87) mm, rotated rx -8.93 ry -0.65 rz 92.62 deg; joints [18.471, 126.68, -173.105, 128.987, 36.186, 117.039, 80.597, 2419.696, 111.51]
  MoveL 26 to (900, 700, 155.68) mm, rotated rx -8.77 ry -1.97 rz 92.59 deg; joints [17.602, 125.932, -173.105, 126.427, 36.839, 119.899, 78.346, 2517.961, 111.514]
  MoveL 27 to (900, 800, 161.12) mm, rotated rx -8.41 ry -3.24 rz 93.06 deg; joints [16.287, 125.726, -173.105, 125.039, 38.529, 122.23, 78.346, 2609.517, 120.738]
  MoveL 28 to (900, 900, 170.13) mm, rotated rx -7.78 ry -6.73 rz 89.38 deg; joints [10.692, 123.529, -173.105, 119.214, 40.759, 128.665, 48.264, 2650.22, 119.321]
  MoveL 29 to (900, 1000, 235.7) mm, rotated rx -45.1 ry -25.31 rz 142.46 deg; joints [-9.5, 123.529, -173.105, 118.036, 88.049, 186.845, 188.236, 2650.23, 426.948]
  Set speed (1000.0 mm/s)
  MoveL 30 to (900, 1000, 235.7) mm, rotated rx -45.1 ry -25.31 rz 142.46 deg; joints [-9.5, 123.529, -173.105, 118.036, 88.049, 186.845, 188.236, 2650.23, 426.948]
  MoveL 31 to (919.24, 1074.55, 171.89) mm, rotated rx -45.1 ry -25.31 rz 142.46 deg; joints [-9.5, 123.529, -173.105, 118.036, 88.05, 186.845, 167.795, 2725.593, 364.48]
  Set speed (1000.0 mm/s)
  MoveL 32 to (838.01, 910.57, 61.58) mm, rotated rx -9.59 ry -1.02 rz 123.08 deg; joints [12.768, 119.824, -159.322, 140.914, 58.982, 136.386, 168.508, 2670.915, 0]
  MoveL 33 to (825, 900, 160.16) mm, rotated rx -9.59 ry -1.02 rz 123.08 deg; joints [12.768, 119.824, -159.322, 140.914, 58.982, 136.386, 183.373, 2659.076, 98.178]
  MoveL 34 to (825, 900, 160.16) mm, rotated rx -8.57 ry 4.45 rz 156.33 deg; joints [17.033, 106.823, -134.821, 156.692, 77.143, 150.504, 183.553, 2659.528, 20.514]
  Set speed (200.0 mm/s)
  MoveL 35 to (825, 800, 150.49) mm, rotated rx -6.95 ry 5.54 rz 156.48 deg; joints [18.123, 106.626, -134.58, 158.309, 76.68, 148.595, 185.525, 2562.17, 2.385]
  MoveL 36 to (825, 700, 144.71) mm, rotated rx -5.29 ry 6.28 rz 156.42 deg; joints [19.27, 106.544, -132.993, 159.782, 77.878, 145.88, 185.526, 2468.907, 0.025]
  MoveL 37 to (825, 600, 141.87) mm, rotated rx -4.02 ry 6.65 rz 156.54 deg; joints [19.969, 106.276, -131.338, 160.87, 79.349, 144.073, 185.528, 2371.682, 0.005]
  MoveL 38 to (825, 500, 141.04) mm, rotated rx -2.81 ry 7.3 rz 156.51 deg; joints [20.71, 106.173, -130.344, 161.988, 80.089, 142.31, 185.528, 2274.13, 0.002]
  MoveL 39 to (825, 400, 142.32) mm, rotated rx -2.04 ry 7.63 rz 156.66 deg; joints [21.668, 106.116, -129.997, 162.549, 80.299, 141.004, 190.959, 2183.637, 0.005]
  MoveL 40 to (825, 300, 145.7) mm, rotated rx -0.73 ry 8.07 rz 156.66 deg; joints [22.115, 105.678, -128.961, 163.631, 81.146, 139.591, 191.811, 2080.761, 0.139]
  MoveL 41 to (825, 200, 151.1) mm, rotated rx 0.43 ry 8.74 rz 156.89 deg; joints [23.404, 105.524, -128.923, 164.564, 80.921, 137.912, 199.843, 1991.049, 0.057]
  MoveL 42 to (825, 100, 159.44) mm, rotated rx 2.11 ry 9.43 rz 156.91 deg; joints [23.984, 104.906, -128.203, 165.984, 81.373, 136.292, 202.469, 1885.88, 0.131]
  MoveL 43 to (825, 0, 171.69) mm, rotated rx 3.99 ry 9.87 rz 156.94 deg; joints [24.453, 103.983, -127.372, 167.342, 82.008, 134.743, 207.291, 1778.17, 1.015]
  Set speed (1000.0 mm/s)
  MoveL 44 to (825, 0, 171.69) mm, rotated rx 3.99 ry 9.87 rz 156.94 deg; joints [24.453, 103.983, -127.372, 167.342, 82.008, 134.743, 207.291, 1778.17, 1.015]
  MoveL 45 to (838.01, -13.11, 73.41) mm, rotated rx 3.99 ry 9.87 rz 156.94 deg; joints [24.453, 105.656, -117.22, 167.443, 93.549, 132.164, 165.245, 1778.693, 0.103]

